(* IEC 61131-3 sources: Industry-PLC-LLM/data/PLCBEAD_repo/PLCBEAD_PLCEmbed-main/PLC-BEAD/Source/PLC_Programs (part 5) *)

(* ---- DT_TO_SDT.ST ---- *)
TYPE oscat_SDT :
STRUCT
	YEAR : INT;
	MONTH : INT;
	DAY : INT;
	WEEKDAY : INT;
	HOUR : INT;
	MINUTE : INT;
	SECOND : INT;
	MS : INT;
END_STRUCT;
END_TYPE

FUNCTION DT_TO_DATE2:UDINT

	VAR_INPUT
		IN :	UDINT;
	END_VAR

	DT_TO_DATE2 := (IN / UDINT#86400) * UDINT#86400;
END_FUNCTION

FUNCTION YEAR_OF_DATE:INT
	VAR_INPUT
		IDATE :	UDINT;
	END_VAR

	YEAR_OF_DATE := UDINT_TO_INT((idate+UDINT#43200) / UDINT#31557600 + UDINT#1970);
END_FUNCTION

FUNCTION DAY_OF_WEEK:INT

	VAR_INPUT
		IDATE :	UDINT;
	END_VAR

	DAY_OF_WEEK := UDINT_TO_INT((idate / UDINT#86400 + UDINT#3) MOD UDINT#7) + INT#01;
END_FUNCTION

FUNCTION LEAP_OF_DATE:BOOL

	VAR_INPUT
		IDATE :	UDINT;
	END_VAR

	LEAP_OF_DATE := SHL(UDINT_TO_DWORD((idate + UDINT#43200) / UDINT#31557600), 30) = DWORD#16#80000000;
END_FUNCTION

FUNCTION DAY_OF_YEAR:INT
	VAR_INPUT
		IDATE :	UDINT;
	END_VAR

	DAY_OF_YEAR := UDINT_TO_INT(((idate) / UDINT#86400) MOD UDINT#1461);
	IF DAY_OF_YEAR > 729 THEN
		IF DAY_OF_YEAR > 1095 THEN DAY_OF_YEAR := DAY_OF_YEAR - 1095; ELSE DAY_OF_YEAR := DAY_OF_YEAR - 729; END_IF;
	ELSIF DAY_OF_YEAR > 364 THEN
		DAY_OF_YEAR := DAY_OF_YEAR - 364;
	ELSE
		DAY_OF_YEAR := DAY_OF_YEAR + 1;
	END_IF;
END_FUNCTION

FUNCTION MONTH_OF_DATE:INT

	VAR_INPUT
		IDATE :	UDINT;
	END_VAR

	MONTH_OF_DATE := DAY_OF_YEAR(idate);
	IF MONTH_OF_DATE < 32 THEN
		MONTH_OF_DATE := 1;
	ELSIF LEAP_OF_DATE((IDATE)) THEN
		MONTH_OF_DATE := (MONTH_OF_DATE * 53 + 1668) / 1623;
	ELSE
		MONTH_OF_DATE := (MONTH_OF_DATE * 53 + 1700) / 1620;
	END_IF;
END_FUNCTION

FUNCTION DAY_OF_MONTH:INT
	VAR_INPUT
		IDATE :	UDINT;
	END_VAR

	day_of_month := day_of_year(idate);

	IF leap_of_Date((idate)) THEN
		CASE day_of_month OF
			32..60	:	day_of_month := day_of_month - 31;
			61..91	:	day_of_month := day_of_month - 60;
			92..121 :	day_of_month := day_of_month - 91;
			122..152:	day_of_month := day_of_month - 121;
			153..182:	day_of_month := day_of_month - 152;
			183..213:	day_of_month := day_of_month - 182;
			214..244:	day_of_month := day_of_month - 213;
			245..274:	day_of_month := day_of_month - 244;
			275..305:	day_of_month := day_of_month - 274;
			306..335:	day_of_month := day_of_month - 305;
			336..366:	day_of_month := day_of_month - 335;
		END_CASE;
	ELSE
		CASE day_of_month OF
			32..59	:	day_of_month := day_of_month - 31;
			60..90	:	day_of_month := day_of_month - 59;
			91..120 :	day_of_month := day_of_month - 90;
			121..151:	day_of_month := day_of_month - 120;
			152..181:	day_of_month := day_of_month - 151;
			182..212:	day_of_month := day_of_month - 181;
			213..243:	day_of_month := day_of_month - 212;
			244..273:	day_of_month := day_of_month - 243;
			274..304:	day_of_month := day_of_month - 273;
			305..334:	day_of_month := day_of_month - 304;
			335..365:	day_of_month := day_of_month - 334;
		END_CASE;
	END_IF;
END_FUNCTION

FUNCTION _INT_TO_UDINT:UDINT
	VAR_INPUT
		IN :	INT;
	END_VAR

	_INT_TO_UDINT := DINT_TO_UDINT(INT_TO_DINT(IN));
END_FUNCTION

FUNCTION_BLOCK DT_TO_SDT

	VAR_INPUT
		DTI :	UDINT;
	END_VAR

	VAR_OUTPUT
		SDT :	oscat_SDT;
	END_VAR

	VAR
		tmp :	UDINT;
		tdt :	UDINT;
	END_VAR

	tmp := DT_TO_DATE2(dti);
	tdt := dti - tmp;
	SDT.YEAR := YEAR_OF_DATE(tmp);
	SDT.MONTH := MONTH_OF_DATE(tmp);
	SDT.DAY := DAY_OF_MONTH(tmp);
	SDT.WEEKDAY := DAY_OF_WEEK(tmp);
	SDT.SECOND := UDINT_TO_INT(tdt MOD UDINT#60);
	SDT.MINUTE := UDINT_TO_INT((tdt / UDINT#60) MOD UDINT#60);
	SDT.HOUR := UDINT_TO_INT(tdt / UDINT#3600);

END_FUNCTION_BLOCK

PROGRAM program0
  VAR
    LocalVar0 : UDINT;
	LocalOUT  : oscat_SDT;
	func_block : DT_TO_SDT;
  END_VAR
	func_block.DTI  := LocalVar0;
	func_block();
	LocalOUT := func_block.SDT;
END_PROGRAM

CONFIGURATION Config0
  RESOURCE Res0 ON PLC
    TASK task0(INTERVAL := T#20ms,PRIORITY := 0);
    PROGRAM instance0 WITH task0 : program0;
  END_RESOURCE
END_CONFIGURATION

(* ---- DT_TO_STRF.ST ---- *)
FUNCTION DT_TO_DATE2:UDINT

	VAR_INPUT
		IN :	UDINT;
	END_VAR

	DT_TO_DATE2 := (IN / UDINT#86400) * UDINT#86400;
END_FUNCTION

FUNCTION DT_TO_TOD2:UDINT
	VAR_INPUT
		IN :	UDINT;
	END_VAR

	DT_TO_TOD2 := (IN MOD UDINT#86400) * UDINT#1000;
END_FUNCTION

FUNCTION _BYTE_TO_INT:INT
	VAR_INPUT
		IN :	BYTE;
	END_VAR

	_BYTE_TO_INT := USINT_TO_INT(BYTE_TO_USINT(IN));
END_FUNCTION

FUNCTION_BLOCK DT_TO_STRF_Block

	VAR_INPUT
		DTI :	UDINT;
		MS :	INT;
		FMT :	STRING;
		LANG :	INT;
	END_VAR

	VAR_OUTPUT
		DT_TO_STRF :	STRING;
	END_VAR

	VAR
		FILL :	STRING;
		BLANK :	STRING;
		ly :	INT;
		dx :	UDINT;
		fs :	STRING;
		fs_tmp :	STRING;
		td :	UDINT;
		tmp :	INT;
		pos :	INT;
		f :	INT;
		CODEE :	CODE;
		MONTH_TO_STRING :	MONTH_TO_STRING;
		WEEKDAY_TO_STRING :	WEEKDAY_TO_STRING;
	END_VAR

	IF LANG < 1 THEN ly := 1; ELSE ly := MIN(2, LANG); END_IF;

	dx := DT_TO_DATE2(DTI);
	td := DT_TO_TOD2(DTI);

	DT_TO_STRF := FMT;
	pos := FIND(DT_TO_STRF, '#');
	WHILE pos > 0 DO
		CODEE(STR:=DT_TO_STRF,POS:=pos + 1);
		f := _BYTE_TO_INT(CODEE.CODEE);
		(* generate the return string according to the format character *)
		fs := '';
		CASE f OF
			0: RETURN; (* illegal character index *)

			65 : (* letter A retunrs the year in 4 digits *)
				fs := INT_TO_STRING(YEAR_OF_DATE(dx),'%d');
			66 : (* letter B returns the year in exactly 2 digits *)
				fs := RIGHT(INT_TO_STRING(YEAR_OF_DATE(dx),'%02d'),2);
			67 : (* letter C returns the month with 1 or 2 digits *)
				fs := INT_TO_STRING(MONTH_OF_DATE(dx),'%d');
			68 : (* letter D returns the month with exactly 2 digits *)
				fs := INT_TO_STRING(MONTH_OF_DATE(dx),'%02d');
			69 : (* letter E returns the month with 3 characters *)
				MONTH_TO_STRING(MTH:=MONTH_OF_DATE(dx),LANG:=ly,LX:=3);
				fs:=MONTH_TO_STRING.MONTH_TO_STRING;
			70 : (* letter F returns the month with all characters *)
				MONTH_TO_STRING(MTH:=MONTH_OF_DATE(dx),LANG:=ly,LX:=0);
				fs:=MONTH_TO_STRING.MONTH_TO_STRING;
			71 : (* letter G returns the day with up to 2 digits *)
				fs := INT_TO_STRING(DAY_OF_MONTH(dx),'%d');
			72 : (* letter H returns the day of the month with exactly 2 digits *)
				fs := INT_TO_STRING(DAY_OF_MONTH(dx),'%d');
				IF LEN(fs) < 2 THEN fs_tmp:=fs; fs := CONCAT(FILL, fs_tmp); END_IF;
			73 : (* letter I returns the weekday as the number 1..7 1 = monday *)
				fs := INT_TO_STRING(DAY_OF_WEEK(dx),'%d');
			74 : (* letter J returns the weekday in 2 character writing *)
				WEEKDAY_TO_STRING(WDAY:=DAY_OF_WEEK(dx),LANG:=ly,LX:=2);
				fs := WEEKDAY_TO_STRING.WEEKDAY_TO_STRING;
			75 : (* letter K returns the weekday with all characters *)
				WEEKDAY_TO_STRING(WDAY:=DAY_OF_WEEK(dx),LANG:=ly,LX:=0);
				fs := WEEKDAY_TO_STRING.WEEKDAY_TO_STRING;
			76 : (* letter L returns AM or PM for the given DateTime *)
				IF td >= UDINT#43200000 THEN fs := 'PM'; ELSE fs := 'AM'; END_IF;
			77 : (* letter M returns the hour in 1 or 2 digit form 0..24h *)
				fs := INT_TO_STRING(HOUR(td),'%d');
			78 : (* letter N returns the hour in exactly 2 digit form 0..24h *)
				fs := INT_TO_STRING(HOUR(td),'%d');
				IF LEN(fs) < 2 THEN fs_tmp:=fs; fs := CONCAT(FILL, fs_tmp); END_IF;
			79 : (* letter O returns the hour in 1 or 2 digit form 0..12h *)
				tmp := HOUR(td) MOD 12;
				IF tmp = 0 THEN tmp := 12; END_IF;
				fs := INT_TO_STRING(tmp,'%d');
			80 : (* letter P returns the hour in exactly 2 digit form 0..12h *)
				tmp := HOUR(td) MOD 12;
				IF tmp = 0 THEN tmp := 12; END_IF;
				fs := INT_TO_STRING(tmp,'%d');
				IF LEN(fs) < 2 THEN fs_tmp:=fs; fs := CONCAT(FILL, fs_tmp); END_IF;
			81 : (* letter Q returns the minute of the hour in 1 or two digit form *)
				fs := INT_TO_STRING(MINUTE(td),'%d');
			82 : (* letter R returns the minute of the hour in exactly two digit form *)
				fs := INT_TO_STRING(MINUTE(td),'%d');
				IF LEN(fs) < 2 THEN fs_tmp:=fs; fs := CONCAT(FILL, fs_tmp); END_IF;
			83 : (* letter S returns the second of the minute in 1 or two digit form *)
				fs := INT_TO_STRING(REAL_TO_INT(SECOND(td)),'%d');
			84 : (* letter T returns the second of the minute in exactly two digit form *)
				fs := INT_TO_STRING(REAL_TO_INT(SECOND(td)),'%d');
				IF LEN(fs) < 2 THEN fs_tmp:=fs; fs := CONCAT(FILL, fs_tmp); END_IF;
			85 : (* letter U returns the milliseconds in 1 to 3 digits *)
				fs := INT_TO_STRING(MS,'%d');
			86 : (* letter V returns the milliseconds in exactly 3 digit form *)
				fs := INT_TO_STRING(MS,'%03d');
			87 : (* letter W returns the day of the month with exactly 2 digits first digit is filled with blank if necessary *)
				fs := INT_TO_STRING(DAY_OF_MONTH(dx),'%d');
				IF LEN(fs) < 2 THEN fs_tmp:=fs; fs := CONCAT(BLANK, fs_tmp); END_IF;
			88 : (* letter X returns the month with exactly 2 digits first digit is filled with blank if necessary *)
				fs := INT_TO_STRING(MONTH_OF_DATE(dx),'%d');
				IF LEN(fs) < 2 THEN fs_tmp:=fs; fs := CONCAT(BLANK, fs_tmp); END_IF;
		END_CASE;
		DT_TO_STRF := REPLACE(DT_TO_STRF, fs, 2, pos);
		pos := FIND(DT_TO_STRF, '#');
	END_WHILE;

END_FUNCTION_BLOCK

PROGRAM program0
  VAR
	DTI  :	UDINT;
	MS   :	INT;
	FMT  :	STRING;
	LANG :	INT;

	DT_TO_STRF :	STRING;

	func_block : DT_TO_STRF_Block;
  END_VAR
	func_block.DTI  :=DTI ;
	func_block.MS   :=MS  ;
	func_block.FMT  :=FMT ;
	func_block.LANG :=LANG;
	func_block();
	DT_TO_STRF := func_block.DT_TO_STRF;
END_PROGRAM

CONFIGURATION Config0
  RESOURCE Res0 ON PLC
    TASK task0(INTERVAL := T#20ms,PRIORITY := 0);
    PROGRAM instance0 WITH task0 : program0;
  END_RESOURCE
END_CONFIGURATION

(* ---- DT_TO_STRING.ST ---- *)
FUNCTION YEAR_OF_DATE:INT
	VAR_INPUT
		IDATE :	UDINT;
	END_VAR

	YEAR_OF_DATE := UDINT_TO_INT((idate+UDINT#43200) / UDINT#31557600 + UDINT#1970);
END_FUNCTION

FUNCTION DAY_OF_YEAR:INT
	VAR_INPUT
		IDATE :	UDINT;
	END_VAR

	DAY_OF_YEAR := UDINT_TO_INT(((idate) / UDINT#86400) MOD UDINT#1461);
	IF DAY_OF_YEAR > 729 THEN
		IF DAY_OF_YEAR > 1095 THEN DAY_OF_YEAR := DAY_OF_YEAR - 1095; ELSE DAY_OF_YEAR := DAY_OF_YEAR - 729; END_IF;
	ELSIF DAY_OF_YEAR > 364 THEN
		DAY_OF_YEAR := DAY_OF_YEAR - 364;
	ELSE
		DAY_OF_YEAR := DAY_OF_YEAR + 1;
	END_IF;
END_FUNCTION

FUNCTION LEAP_OF_DATE:BOOL

	VAR_INPUT
		IDATE :	UDINT;
	END_VAR

	LEAP_OF_DATE := SHL(UDINT_TO_DWORD((idate + UDINT#43200) / UDINT#31557600), 30) = DWORD#16#80000000;
END_FUNCTION

FUNCTION MONTH_OF_DATE:INT

	VAR_INPUT
		IDATE :	UDINT;
	END_VAR

	MONTH_OF_DATE := DAY_OF_YEAR(idate);
	IF MONTH_OF_DATE < 32 THEN
		MONTH_OF_DATE := 1;
	ELSIF LEAP_OF_DATE(IDATE) THEN
		MONTH_OF_DATE := (MONTH_OF_DATE * 53 + 1668) / 1623;
	ELSE
		MONTH_OF_DATE := (MONTH_OF_DATE * 53 + 1700) / 1620;
	END_IF;
END_FUNCTION

FUNCTION DAY_OF_MONTH:INT
	VAR_INPUT
		IDATE :	UDINT;
	END_VAR

	day_of_month := day_of_year(idate);

	IF leap_of_Date((idate)) THEN
		CASE day_of_month OF
			32..60	:	day_of_month := day_of_month - 31;
			61..91	:	day_of_month := day_of_month - 60;
			92..121 :	day_of_month := day_of_month - 91;
			122..152:	day_of_month := day_of_month - 121;
			153..182:	day_of_month := day_of_month - 152;
			183..213:	day_of_month := day_of_month - 182;
			214..244:	day_of_month := day_of_month - 213;
			245..274:	day_of_month := day_of_month - 244;
			275..305:	day_of_month := day_of_month - 274;
			306..335:	day_of_month := day_of_month - 305;
			336..366:	day_of_month := day_of_month - 335;
		END_CASE;
	ELSE
		CASE day_of_month OF
			32..59	:	day_of_month := day_of_month - 31;
			60..90	:	day_of_month := day_of_month - 59;
			91..120 :	day_of_month := day_of_month - 90;
			121..151:	day_of_month := day_of_month - 120;
			152..181:	day_of_month := day_of_month - 151;
			182..212:	day_of_month := day_of_month - 181;
			213..243:	day_of_month := day_of_month - 212;
			244..273:	day_of_month := day_of_month - 243;
			274..304:	day_of_month := day_of_month - 273;
			305..334:	day_of_month := day_of_month - 304;
			335..365:	day_of_month := day_of_month - 334;
		END_CASE;
	END_IF;
END_FUNCTION

FUNCTION SECOND_OF_DT:INT

	VAR_INPUT
		XDT :	UDINT;
	END_VAR

	SECOND_OF_DT := UDINT_TO_INT(XDT MOD UDINT#60);
END_FUNCTION

FUNCTION HOUR_OF_DT:INT
	VAR_INPUT
		XDT :	UDINT;
	END_VAR

	HOUR_OF_DT := UDINT_TO_INT((XDT MOD UDINT#86400) / UDINT#3600);
END_FUNCTION

FUNCTION MINUTE_OF_DT:INT
	VAR_INPUT
		XDT :	UDINT;
	END_VAR

	MINUTE_OF_DT := UDINT_TO_INT((XDT MOD UDINT#3600) / UDINT#60);
END_FUNCTION

FUNCTION_BLOCK DT_TO_STRING_Block

	VAR_INPUT
		IDT :	UDINT;
	END_VAR

	VAR_OUTPUT
		DT_STRING :	STRING;
	END_VAR

	VAR
		st_tmp1 :	STRING;
		st_tmp2 :	STRING;
	END_VAR

	st_tmp2 := CONCAT(INT_TO_STRING(YEAR_OF_DATE(IDT)),INT_TO_STRING(MONTH_OF_DATE(IDT)));
	st_tmp1 := CONCAT(INT_TO_STRING(day_of_month(IDT)),INT_TO_STRING(hour_of_DT(IDT)));
	st_tmp2 := CONCAT(st_tmp2,st_tmp1);
	st_tmp1 := CONCAT(INT_TO_STRING(minute_of_DT(IDT)),INT_TO_STRING(second_of_DT(IDT)));
	st_tmp2 := CONCAT(st_tmp2,st_tmp1);
	DT_STRING := st_tmp2;
END_FUNCTION_BLOCK

PROGRAM program0
	VAR
		IDT : UDINT;
		OUT  : STRING;
		func_block : DT_TO_STRING_Block;
	END_VAR
	func_block.IDT := IDT;
	func_block();
	OUT := func_block.DT_STRING;
END_PROGRAM

CONFIGURATION Config0
	RESOURCE Res0 ON PLC
		TASK task0(INTERVAL := T#20ms,PRIORITY := 0);
		PROGRAM instance0 WITH task0 : program0;
	END_RESOURCE
END_CONFIGURATION

(* ---- DW_TO_REAL.ST ---- *)
FUNCTION_BLOCK DW_TO_REAL_Block
  VAR_INPUT
    X :	DWORD;
  END_VAR

  VAR_OUTPUT
    DW_TO_REAL :	REAL;
  END_VAR

  VAR
    BUF_TO_REAL :	BUF_TO_REAL;
    i :	INT;
  END_VAR

  FOR I := 0 TO 1 DO
    BUF_TO_REAL.REQ        := I > 0;
    BUF_TO_REAL.BUF_FORMAT := FALSE;
    BUF_TO_REAL.BUF_OFFS   := DINT#0;
    BUF_TO_REAL.BUF_CNT    := DINT#4;
    BUF_TO_REAL.BUFFER     := X;
    BUF_TO_REAL.DST        := DW_TO_REAL;
    BUF_TO_REAL();
    X           := BUF_TO_REAL.BUFFER;
    DW_TO_REAL  := BUF_TO_REAL.DST;
  END_FOR;
END_FUNCTION_BLOCK

(* ---- DWORD_TO_STRB.ST ---- *)
FUNCTION_BLOCK DWORD_TO_STRB_Block
	VAR_INPUT
		IN :	DWORD;
	END_VAR

	VAR_OUTPUT
		DWORD_TO_STRB :	STRING;
	END_VAR

	VAR
		i :	INT;
	END_VAR

	DWORD_TO_STRB :='';
	FOR i := 1 TO 32 DO
		IF (in AND DWORD#16#8000_0000) > DWORD#0 THEN
			DWORD_TO_STRB := CONCAT(DWORD_TO_STRB,'1');
		ELSE
			DWORD_TO_STRB := CONCAT(DWORD_TO_STRB,'0');
		END_IF;
		in := SHL(in, 1);
	END_FOR;
END_FUNCTION_BLOCK

PROGRAM program0
  VAR
    IN :	DWORD;

	DWORD_TO_STRB :	STRING;
	func_block : DWORD_TO_STRB_Block;
  END_VAR
	func_block.IN  := IN;
	func_block();
	DWORD_TO_STRB := func_block.DWORD_TO_STRB;
END_PROGRAM

CONFIGURATION Config0
  RESOURCE Res0 ON PLC
    TASK task0(INTERVAL := T#20ms,PRIORITY := 0);
    PROGRAM instance0 WITH task0 : program0;
  END_RESOURCE
END_CONFIGURATION

(* ---- DWORD_TO_STRF.ST ---- *)
FUNCTION_BLOCK DWORD_TO_STRF_Block

	VAR_INPUT
		IN :	DWORD;
		N :	INT;
	END_VAR

	VAR_OUTPUT
		DWORD_TO_STRF :	STRING;
	END_VAR

	VAR
		temp :	STRING;
		temp2 :	STRING;
		L : INT;
	END_VAR

	temp := DWORD_TO_STRING(in);
	L := LEN(temp);
	IF N < L THEN
		temp :=RIGHT(temp,N);
		L := N;
	END_IF;

	WHILE L < N DO
		temp2 := temp;
		temp := CONCAT('0', temp2);
		L := L + 1;
	END_WHILE;
	DWORD_TO_STRF := temp;

END_FUNCTION_BLOCK

PROGRAM program0
  VAR
    IN :	DWORD;
	N :		INT;
	DWORD_TO_STRF :	STRING;
	func_block : DWORD_TO_STRF_Block;
  END_VAR
	func_block.IN  := IN;
	func_block.N  := N;
	func_block();
	DWORD_TO_STRF := func_block.DWORD_TO_STRF;
END_PROGRAM

CONFIGURATION Config0
  RESOURCE Res0 ON PLC
    TASK task0(INTERVAL := T#20ms,PRIORITY := 0);
    PROGRAM instance0 WITH task0 : program0;
  END_RESOURCE
END_CONFIGURATION

(* ---- DWORD_TO_STRH.ST ---- *)
FUNCTION_BLOCK DWORD_TO_STRH_Block

	VAR_INPUT
		IN :	DWORD;
	END_VAR

	VAR_OUTPUT
		DWORD_TO_STRH :	STRING;
	END_VAR

	DWORD_TO_STRH:=DWORD_TO_STRING(IN);

END_FUNCTION_BLOCK

PROGRAM program0
  VAR
    LocalVar0 : DWORD;
	LocalOUT  : STRING;
	func_block : DWORD_TO_STRH_Block;
  END_VAR
	func_block.IN  := LocalVar0;
	func_block();
	LocalOUT := func_block.DWORD_TO_STRH;
END_PROGRAM

CONFIGURATION Config0
  RESOURCE Res0 ON PLC
    TASK task0(INTERVAL := T#20ms,PRIORITY := 0);
    PROGRAM instance0 WITH task0 : program0;
  END_RESOURCE
END_CONFIGURATION

(* ---- ELEMENT_COUNT.ST ---- *)
TYPE
	oscat_STRING250             : STRING;
END_TYPE

FUNCTION_BLOCK ELEMENT_COUNT_Block

	VAR_IN_OUT
		ELEMENT :	oscat_STRING250;
	END_VAR

	VAR_INPUT
		SEP :	BYTE;
	END_VAR

	VAR_OUTPUT
		ELEMENT_COUNT :	INT;
	END_VAR

	VAR
		I :	INT;
		pos :	INT;
	END_VAR

	i := LEN(ELEMENT);
	IF i = 0 THEN
		ELEMENT_COUNT := 0;
	ELSE
		ELEMENT_COUNT := 1;
		FOR pos := 1 TO I DO
			IF INT_TO_BYTE(GET_CHAR(ELEMENT,pos)) = SEP THEN ELEMENT_COUNT := ELEMENT_COUNT + 1; END_IF;
		END_FOR;
	END_IF;

END_FUNCTION_BLOCK

PROGRAM program0
	VAR
		SEP :	BYTE;
		POS :	INT;
		ELEMENT :	oscat_STRING250;
		ELEMENT_GET :	oscat_STRING250;

		func_block : ELEMENT_COUNT_Block;
	END_VAR
	func_block.SEP    :=SEP    ;
	func_block.POS:=POS;
	func_block.ELEMENT     :=ELEMENT     ;
	func_block();
	ELEMENT    := func_block.ELEMENT    ;
	ELEMENT_GET:= func_block.ELEMENT_GET;

END_PROGRAM

CONFIGURATION Config0
  RESOURCE Res0 ON PLC
    TASK task0(INTERVAL := T#20ms,PRIORITY := 0);
    PROGRAM instance0 WITH task0 : program0;
  END_RESOURCE
END_CONFIGURATION

(* ---- ELEMENT_GET.ST ---- *)
TYPE
	oscat_STRING250             : STRING;
END_TYPE

FUNCTION_BLOCK ELEMENT_GET_Block

	VAR_INPUT
		SEP :	BYTE;
		POS :	INT;
	END_VAR

	VAR_IN_OUT
		ELEMENT :	oscat_STRING250;
	END_VAR

	VAR_OUTPUT
		ELEMENT_GET :	oscat_STRING250;
	END_VAR

	VAR
		i :	INT;
		i2 :	INT;
		cnt :	INT;
		size :	INT;
	END_VAR

	cnt := 0;
	size := LEN(ELEMENT);

	FOR i := 1 TO size DO
		IF cnt = POS THEN EXIT; END_IF;
		IF INT_TO_BYTE(GET_CHAR(ELEMENT,i)) = SEP THEN cnt := cnt + 1; END_IF;
	END_FOR;

	FOR i2 := i TO size DO
		IF INT_TO_BYTE(GET_CHAR(ELEMENT,i2)) = SEP THEN EXIT; END_IF;
	END_FOR;

	IF i2 > i THEN
		ELEMENT_GET := MID(ELEMENT,i2-i,i);
	ELSE
		ELEMENT_GET := '';
	END_IF;

END_FUNCTION_BLOCK

PROGRAM program0
	VAR
		SEP :	BYTE;
		POS :	INT;
		ELEMENT :	oscat_STRING250;
		ELEMENT_GET :	oscat_STRING250;

		func_block : ELEMENT_GET_Block;
	END_VAR
	func_block.SEP    :=SEP    ;
	func_block.POS:=POS;
	func_block.ELEMENT     :=ELEMENT     ;
	func_block();
	ELEMENT    := func_block.ELEMENT    ;
	ELEMENT_GET:= func_block.ELEMENT_GET;

END_PROGRAM

CONFIGURATION Config0
  RESOURCE Res0 ON PLC
    TASK task0(INTERVAL := T#20ms,PRIORITY := 0);
    PROGRAM instance0 WITH task0 : program0;
  END_RESOURCE
END_CONFIGURATION

(* ---- ENERGY.ST ---- *)
FUNCTION_BLOCK ENERGY
	VAR_INPUT
		J :	REAL;
		C :	REAL;
		WH :	REAL;
	END_VAR

	VAR_OUTPUT
		YJ :	REAL;
		YC :	REAL;
		YWH :	REAL;
	END_VAR

	YJ := J + Wh * 3600.0 + C * 4.1868;
	YC := YJ * 0.238845896627496;
	YWh := YJ * 2.7777777778E-004;
END_FUNCTION_BLOCK

PROGRAM program0
  VAR
		J  :	REAL;
		C  :	REAL;
		WH :	REAL;

		YJ  :	REAL;
		YC  :	REAL;
		YWH :	REAL;
	func_block : ENERGY;
  END_VAR
	func_block.J  :=J ;
	func_block.C  :=C ;
	func_block.WH :=WH;
	func_block();
	YJ  := func_block.YJ ;
	YC  := func_block.YC ;
	YWH := func_block.YWH;

END_PROGRAM

CONFIGURATION Config0
	RESOURCE Res0 ON PLC
		TASK task0(INTERVAL := T#20ms,PRIORITY := 0);
		PROGRAM instance0 WITH task0 : program0;
	END_RESOURCE
END_CONFIGURATION

(* ---- ESR_COLLECT.ST ---- *)
TYPE
	oscat_esr_collect_data      : ARRAY [0..7]    OF BYTE;
END_TYPE
TYPE oscat_esr_data :
  STRUCT
	typ    : BYTE;
	adress : STRING;
	DS     : UDINT;
	TS     : TIME;
	data   : oscat_esr_collect_data;
  END_STRUCT;
END_TYPE

TYPE
  oscat_ESR_3                : ARRAY [0..3] OF oscat_esr_data;
  oscat_ESR_31               : ARRAY [0..31] OF oscat_esr_data;
END_TYPE

FUNCTION INC1:INT

	VAR_INPUT
		X :	INT;
		N :	INT;
	END_VAR

	IF X >= N - 1 THEN
		INC1 := 0;
	ELSE
		INC1 := X + 1;
	END_IF;
END_FUNCTION

FUNCTION_BLOCK ESR_COLLECT
	VAR_INPUT
		ESR_0 :	oscat_ESR_3;
		ESR_1 :	oscat_ESR_3;
		ESR_2 :	oscat_ESR_3;
		ESR_3 :	oscat_ESR_3;
		ESR_4 :	oscat_ESR_3;
		ESR_5 :	oscat_ESR_3;
		ESR_6 :	oscat_ESR_3;
		ESR_7 :	oscat_ESR_3;
		RST :	BOOL;
	END_VAR

	VAR_IN_OUT
		POS :	INT;
	END_VAR

	VAR_OUTPUT
		ESR_OUT :	oscat_ESR_31;
	END_VAR

	VAR
		cnt :	INT := -1;
		max_in :	INT := 3;
		max_out :	INT := 32;
	END_VAR

	IF rst OR cnt < 0 THEN
		pos := -1;
	ELSE
		FOR cnt := 0 TO max_in DO
		IF esr_0[cnt].typ > BYTE#0 THEN pos := INC1(pos, max_out); esr_out[pos] := esr_0[cnt]; END_IF;
		IF esr_1[cnt].typ > BYTE#0 THEN pos := INC1(pos, max_out); esr_out[pos] := esr_1[cnt]; END_IF;
		IF esr_2[cnt].typ > BYTE#0 THEN pos := INC1(pos, max_out); esr_out[pos] := esr_2[cnt]; END_IF;
		IF esr_3[cnt].typ > BYTE#0 THEN pos := INC1(pos, max_out); esr_out[pos] := esr_3[cnt]; END_IF;
		IF esr_4[cnt].typ > BYTE#0 THEN pos := INC1(pos, max_out); esr_out[pos] := esr_4[cnt]; END_IF;
		IF esr_5[cnt].typ > BYTE#0 THEN pos := INC1(pos, max_out); esr_out[pos] := esr_5[cnt]; END_IF;
		IF esr_6[cnt].typ > BYTE#0 THEN pos := INC1(pos, max_out); esr_out[pos] := esr_6[cnt]; END_IF;
		IF esr_7[cnt].typ > BYTE#0 THEN pos := INC1(pos, max_out); esr_out[pos] := esr_7[cnt]; END_IF;
	END_FOR;
	END_IF;

END_FUNCTION_BLOCK

PROGRAM program0
  VAR
	ESR_0 :	oscat_ESR_3;
	ESR_1 :	oscat_ESR_3;
	ESR_2 :	oscat_ESR_3;
	ESR_3 :	oscat_ESR_3;
	ESR_4 :	oscat_ESR_3;
	ESR_5 :	oscat_ESR_3;
	ESR_6 :	oscat_ESR_3;
	ESR_7 :	oscat_ESR_3;
	RST   :	BOOL;

	POS   :	INT;

	ESR_OUT :	oscat_ESR_31;

	func_block : ESR_COLLECT;
  END_VAR
	func_block.ESR_0 :=ESR_0;
	func_block.ESR_1 :=ESR_1;
	func_block.ESR_2 :=ESR_2;
	func_block.ESR_3 :=ESR_3;
	func_block.ESR_4 :=ESR_4;
	func_block.ESR_5 :=ESR_5;
	func_block.ESR_6 :=ESR_6;
	func_block.ESR_7 :=ESR_7;
	func_block.RST   :=RST  ;
	func_block.POS   :=POS  ;

	func_block();
	POS := func_block.POS;
	ESR_OUT := func_block.ESR_OUT;

END_PROGRAM

CONFIGURATION Config0
	RESOURCE Res0 ON PLC
		TASK task0(INTERVAL := T#20ms,PRIORITY := 0);
		PROGRAM instance0 WITH task0 : program0;
	END_RESOURCE
END_CONFIGURATION

(* ---- ESR_MON_B8.ST ---- *)
TYPE
	oscat_esr_collect_data      : ARRAY [0..7]    OF BYTE;
END_TYPE
TYPE oscat_esr_data :
  STRUCT
	typ    : BYTE;
	adress : STRING;
	DS     : UDINT;
	TS     : TIME;
	data   : oscat_esr_collect_data;
  END_STRUCT;
END_TYPE

TYPE
  oscat_ESR_3                : ARRAY [0..3] OF oscat_esr_data;
  oscat_ESR_31               : ARRAY [0..31] OF oscat_esr_data;
END_TYPE

FUNCTION_BLOCK T_PLC_MS_block

	VAR_OUTPUT
		T_PLC_MS :	UDINT;
	END_VAR

	VAR_EXTERNAL
		PLC_TICKS_PER_SEC :	INT;
		PLC_SYS_TICK_CNT :	DINT;
	END_VAR

	VAR
		debug :	BOOL;(*Debug-Mode ON / OFF*)
		N :	INT;(*Debug-Faktor*)
		Offset :	UDINT;(*Debug-Offset*)
		temp :	DWORD := DWORD#1;(*Debug-Offset*)
		mode :	BOOL;(*modus*)
		faktor :	UDINT;(*Systemtakt-Faktor*)
		init :	BOOL;
		v_plc_ticks_per_sec :	UDINT;
		base :	UDINT := UDINT#1000;
	END_VAR

	IF init = FALSE THEN
		v_plc_ticks_per_sec := INT_TO_UDINT(PLC_TICKS_PER_SEC);
		IF v_plc_ticks_per_sec = UDINT#1024 THEN
			faktor := UDINT#1;
			mode := FALSE;
		ELSIF v_plc_ticks_per_sec > UDINT#0 THEN
			IF v_plc_ticks_per_sec <= base THEN
				faktor := base / v_plc_ticks_per_sec;
				mode := FALSE;
			ELSE
				faktor := v_plc_ticks_per_sec / base;
				mode := TRUE;
			END_IF;
		ELSE
			faktor := UDINT#1;
		END_IF;
		init := TRUE;
	END_IF;

	IF mode THEN
		T_PLC_MS := DINT_TO_UDINT(PLC_SYS_TICK_CNT) / faktor;
	ELSE
		T_PLC_MS := DINT_TO_UDINT(PLC_SYS_TICK_CNT) * faktor;
	END_IF;

	IF debug THEN
		T_PLC_MS := (DWORD_TO_UDINT(SHL(UDINT_TO_DWORD(T_PLC_MS),N) OR SHL(temp,N)) - UDINT#1) + Offset;
	END_IF;

END_FUNCTION_BLOCK

FUNCTION_BLOCK ESR_MON_B8

	VAR_INPUT
		S0 :	BOOL;
		A0 :	STRING;
		S1 :	BOOL;
		A1 :	STRING;
		S2 :	BOOL;
		A2 :	STRING;
		S3 :	BOOL;
		A3 :	STRING;
		S4 :	BOOL;
		A4 :	STRING;
		S5 :	BOOL;
		A5 :	STRING;
		S6 :	BOOL;
		A6 :	STRING;
		S7 :	BOOL;
		A7 :	STRING;
		DT_IN :	UDINT;
	END_VAR

	VAR_IN_OUT
		ESR_Out :	oscat_ESR_3;
	END_VAR

	VAR_OUTPUT
		ESR_FLAG :	BOOL;
	END_VAR

	VAR
		x0 :	BOOL;
		x1 :	BOOL;
		x2 :	BOOL;
		x3 :	BOOL;
		x4 :	BOOL;
		x5 :	BOOL;
		x6 :	BOOL;
		x7 :	BOOL;
		tx :	TIME;
		cnt :	INT;
		T_PLC_MS :	T_PLC_MS_block;
	END_VAR

	T_PLC_MS();
	tx:= UDINT_TO_TIME(T_PLC_MS.T_PLC_MS);

	ESR_Flag := FALSE;
	esr_out[3].typ := BYTE#0;
	esr_out[2].typ := BYTE#0;
	esr_out[1].typ := BYTE#0;
	esr_out[0].typ := BYTE#0;
	cnt := 0;

	IF s0 <> X0 THEN
		esr_out[cnt].typ := INT_TO_BYTE(10 + BOOL_TO_INT(s0));
		esr_out[cnt].adress := a0;
		esr_out[cnt].DS := DT_in;
		esr_out[cnt].TS := TX;
		X0 := S0;
		cnt := cnt + 1;
		esr_flag := TRUE;
	END_IF;
	IF s1 <> X1 THEN
		esr_out[cnt].typ := INT_TO_BYTE(10 + BOOL_TO_INT(s1));
		esr_out[cnt].adress := a1;
		esr_out[cnt].DS := DT_in;
		esr_out[cnt].TS := TX;
		X1 := S1;
		cnt := cnt + 1;
		esr_flag := TRUE;
	END_IF;
	IF s2 <> X2 THEN
		esr_out[cnt].typ := INT_TO_BYTE(10 + BOOL_TO_INT(s2));
		esr_out[cnt].adress := a2;
		esr_out[cnt].DS := DT_in;
		esr_out[cnt].TS := TX;
		X2 := S2;
		cnt := cnt + 1;
		esr_flag := TRUE;
	END_IF;
	IF s3 <> X3 THEN
		esr_out[cnt].typ := INT_TO_BYTE(10 + BOOL_TO_INT(s3));
		esr_out[cnt].adress := a3;
		esr_out[cnt].DS := DT_in;
		esr_out[cnt].TS := TX;
		X3 := S3;
		cnt := cnt + 1;
		esr_flag := TRUE;
	END_IF;
	IF s4 <> X4 AND cnt < 4 THEN
		esr_out[cnt].typ := INT_TO_BYTE(10 + BOOL_TO_INT(s4));
		esr_out[cnt].adress := a4;
		esr_out[cnt].DS := DT_in;
		esr_out[cnt].TS := TX;
		X4 := S4;
		cnt := cnt + 1;
		esr_flag := TRUE;
	END_IF;
	IF s5 <> X5  AND cnt < 4 THEN
		esr_out[cnt].typ := INT_TO_BYTE(10 + BOOL_TO_INT(s5));
		esr_out[cnt].adress := a5;
		esr_out[cnt].DS := DT_in;
		esr_out[cnt].TS := TX;
		X5 := S5;
		cnt := cnt + 1;
		esr_flag := TRUE;
	END_IF;
	IF s6 <> X6  AND cnt < 4 THEN
		esr_out[cnt].typ := INT_TO_BYTE(10 + BOOL_TO_INT(s6));
		esr_out[cnt].adress := a6;
		esr_out[cnt].DS := DT_in;
		esr_out[cnt].TS := TX;
		X6 := S6;
		cnt := cnt + 1;
		esr_flag := TRUE;
	END_IF;
	IF s7 <> X7  AND cnt < 4 THEN
		esr_out[cnt].typ := INT_TO_BYTE(10 + BOOL_TO_INT(s7));
		esr_out[cnt].adress := a7;
		esr_out[cnt].DS := DT_in;
		esr_out[cnt].TS := TX;
		X7 := S7;
		cnt := cnt + 1;
		esr_flag := TRUE;
	END_IF;

END_FUNCTION_BLOCK

PROGRAM program0

	VAR

		S0 :	BOOL;
		A0 :	STRING;
		S1 :	BOOL;
		A1 :	STRING;
		S2 :	BOOL;
		A2 :	STRING;
		S3 :	BOOL;
		A3 :	STRING;
		S4 :	BOOL;
		A4 :	STRING;
		S5 :	BOOL;
		A5 :	STRING;
		S6 :	BOOL;
		A6 :	STRING;
		S7 :	BOOL;
		A7 :	STRING;
		DT_IN   :	UDINT;

		ESR_Out :	oscat_ESR_3;

		ESR_FLAG :	BOOL;

		func_block : ESR_MON_B8;
  	END_VAR
	func_block.S0 := S0;
	func_block.A0 := A0;
	func_block.S1 := S1;
	func_block.A1 := A1;
	func_block.S2 := S2;
	func_block.A2 := A2;
	func_block.S3 := S3;
	func_block.A3 := A3;
	func_block.S4 := S4;
	func_block.A4 := A4;
	func_block.S5 := S5;
	func_block.A5 := A5;
	func_block.S6 := S6;
	func_block.A6 := A6;
	func_block.S7 := S7;
	func_block.A7 := A7;
	func_block.DT_IN := DT_IN;
	func_block.ESR_Out := ESR_Out;
	func_block();
	ESR_Out := func_block.ESR_Out;
	ESR_FLAG := func_block.ESR_FLAG;

END_PROGRAM

CONFIGURATION Config0

	VAR_GLOBAL
		PLC_TICKS_PER_SEC :	INT;
		PLC_SYS_TICK_CNT :	DINT;
	END_VAR

  	RESOURCE Res0 ON PLC
    	TASK task0(INTERVAL := T#20ms,PRIORITY := 0);
    	PROGRAM instance0 WITH task0 : program0;
  	END_RESOURCE

END_CONFIGURATION

(* ---- ESR_MON_R4.ST ---- *)
TYPE
	oscat_esr_collect_data      : ARRAY [0..7]    OF BYTE;
END_TYPE

TYPE oscat_esr_data :
  STRUCT
	typ    : BYTE;
	adress : STRING;
	DS     : UDINT;
	TS     : TIME;
	data   : oscat_esr_collect_data;
  END_STRUCT;
END_TYPE

TYPE
  oscat_ESR_3                : ARRAY [0..3] OF oscat_esr_data;
  oscat_ESR_31               : ARRAY [0..31] OF oscat_esr_data;
END_TYPE

FUNCTION_BLOCK REAL_TO_DW_Block
  VAR_INPUT
    X :	REAL;
  END_VAR

  VAR_OUTPUT
    REAL_TO_DW :	DWORD;
  END_VAR

  VAR
    REAL_TO_BUF :	REAL_TO_BUF;
    i :	INT;
  END_VAR

  FOR I := 0 TO 1 DO
    REAL_TO_BUF.REQ        := I > 0;
    REAL_TO_BUF.BUF_FORMAT := FALSE;
    REAL_TO_BUF.BUF_OFFS   := DINT#0;
    REAL_TO_BUF.BUF_CNT    := DINT#4;
    REAL_TO_BUF.SRC        := X;
    REAL_TO_BUF.BUFFER     := REAL_TO_DW;
    REAL_TO_BUF();
    X          := REAL_TO_BUF.SRC;
    REAL_TO_DW := REAL_TO_BUF.BUFFER;
  END_FOR;
END_FUNCTION_BLOCK

FUNCTION_BLOCK T_PLC_MS_block

	VAR_OUTPUT
		T_PLC_MS :	UDINT;
	END_VAR

	VAR_EXTERNAL
		PLC_TICKS_PER_SEC :	INT;
		PLC_SYS_TICK_CNT :	DINT;
	END_VAR

	VAR
		debug :	BOOL;(*Debug-Mode ON / OFF*)
		N :	INT;(*Debug-Faktor*)
		Offset :	UDINT;(*Debug-Offset*)
		temp :	DWORD := DWORD#1;(*Debug-Offset*)
		mode :	BOOL;(*modus*)
		faktor :	UDINT;(*Systemtakt-Faktor*)
		init :	BOOL;
		v_plc_ticks_per_sec :	UDINT;
		base :	UDINT := UDINT#1000;
	END_VAR

	IF init = FALSE THEN
		v_plc_ticks_per_sec := INT_TO_UDINT(PLC_TICKS_PER_SEC);
		IF v_plc_ticks_per_sec = UDINT#1024 THEN
			faktor := UDINT#1;
			mode := FALSE;
		ELSIF v_plc_ticks_per_sec > UDINT#0 THEN
			IF v_plc_ticks_per_sec <= base THEN
				faktor := base / v_plc_ticks_per_sec;
				mode := FALSE;
			ELSE
				faktor := v_plc_ticks_per_sec / base;
				mode := TRUE;
			END_IF;
		ELSE
			faktor := UDINT#1;
		END_IF;
		init := TRUE;
	END_IF;

	IF mode THEN
		T_PLC_MS := DINT_TO_UDINT(PLC_SYS_TICK_CNT) / faktor;
	ELSE
		T_PLC_MS := DINT_TO_UDINT(PLC_SYS_TICK_CNT) * faktor;
	END_IF;

	IF debug THEN
		T_PLC_MS := (DWORD_TO_UDINT(SHL(UDINT_TO_DWORD(T_PLC_MS),N) OR SHL(temp,N)) - UDINT#1) + Offset;
	END_IF;

END_FUNCTION_BLOCK

FUNCTION_BLOCK ESR_MON_R4
	VAR_INPUT
		R0 :	REAL;
		A0 :	STRING;
		S0 :	REAL;
		R1 :	REAL;
		A1 :	STRING;
		S1 :	REAL;
		R2 :	REAL;
		A2 :	STRING;
		S2 :	REAL;
		R3 :	REAL;
		A3 :	STRING;
		S3 :	REAL;
		DT_IN :	UDINT;
	END_VAR

	VAR_IN_OUT
		ESR_OUT :	oscat_ESR_3;
	END_VAR

	VAR_OUTPUT
		ESR_FLAG :	BOOL;
	END_VAR

	VAR
		x0 :	REAL;
		x1 :	REAL;
		x2 :	REAL;
		x3 :	REAL;
		tx :	TIME;
		cnt :	INT;
		T_PLC_MS :	T_PLC_MS_block;
		REAL_TO_DW :	REAL_TO_DW_Block;
		tmp :	DWORD;
	END_VAR

	T_PLC_MS();
	tx:= UDINT_TO_TIME(T_PLC_MS.T_PLC_MS);

	ESR_Flag := FALSE;
	esr_out[3].typ := BYTE#0;
	esr_out[2].typ := BYTE#0;
	esr_out[1].typ := BYTE#0;
	esr_out[0].typ := BYTE#0;
	cnt := 0;

	IF differ(R0, X0, S0) THEN
		REAL_TO_DW(X:=R0);
		tmp := REAL_TO_DW.REAL_TO_DW;

		esr_out[cnt].typ := BYTE#20;
		esr_out[cnt].adress := a0;
		esr_out[cnt].DS := DT_in;
		esr_out[cnt].TS := TX;
		esr_out[cnt].data[0] := Byte_of_Dword(tmp,BYTE#0);
		esr_out[cnt].data[1] := Byte_of_Dword(tmp,BYTE#1);
		esr_out[cnt].data[2] := Byte_of_Dword(tmp,BYTE#2);
		esr_out[cnt].data[3] := Byte_of_Dword(tmp,BYTE#3);
		X0 := R0;
		cnt := cnt + 1;
		esr_flag := TRUE;
	END_IF;
	IF differ(R1, X1, S1) THEN
		REAL_TO_DW(X:=R1);
		tmp := REAL_TO_DW.REAL_TO_DW;

		esr_out[cnt].typ := BYTE#20;
		esr_out[cnt].adress := a1;
		esr_out[cnt].DS := DT_in;
		esr_out[cnt].TS := TX;
		esr_out[cnt].data[0] := Byte_of_Dword(tmp,BYTE#0);
		esr_out[cnt].data[1] := Byte_of_Dword(tmp,BYTE#1);
		esr_out[cnt].data[2] := Byte_of_Dword(tmp,BYTE#2);
		esr_out[cnt].data[3] := Byte_of_Dword(tmp,BYTE#3);
		X1 := R1;
		cnt := cnt + 1;
		esr_flag := TRUE;
	END_IF;
	IF differ(R2, X2, S2) THEN
		REAL_TO_DW(X:=R2);
		tmp := REAL_TO_DW.REAL_TO_DW;

		esr_out[cnt].typ := BYTE#20;
		esr_out[cnt].adress := a2;
		esr_out[cnt].DS := DT_in;
		esr_out[cnt].TS := TX;
		esr_out[cnt].data[0] := Byte_of_Dword(tmp,BYTE#0);
		esr_out[cnt].data[1] := Byte_of_Dword(tmp,BYTE#1);
		esr_out[cnt].data[2] := Byte_of_Dword(tmp,BYTE#2);
		esr_out[cnt].data[3] := Byte_of_Dword(tmp,BYTE#3);
		X2 := R2;
		cnt := cnt + 1;
		esr_flag := TRUE;
	END_IF;
	IF differ(R3, X3, S3) THEN
		REAL_TO_DW(X:=R2);
		tmp := REAL_TO_DW.REAL_TO_DW;

		esr_out[cnt].typ := BYTE#20;
		esr_out[cnt].adress := a3;
		esr_out[cnt].DS := DT_in;
		esr_out[cnt].TS := TX;
		esr_out[cnt].data[0] := Byte_of_Dword(tmp,BYTE#0);
		esr_out[cnt].data[1] := Byte_of_Dword(tmp,BYTE#1);
		esr_out[cnt].data[2] := Byte_of_Dword(tmp,BYTE#2);
		esr_out[cnt].data[3] := Byte_of_Dword(tmp,BYTE#3);
		X3 := R3;
		cnt := cnt + 1;
		esr_flag := TRUE;
	END_IF;
END_FUNCTION_BLOCK

PROGRAM program0

	VAR
	VAR_INPUT
		R0 :	REAL;
		A0 :	STRING;
		S0 :	REAL;
		R1 :	REAL;
		A1 :	STRING;
		S1 :	REAL;
		R2 :	REAL;
		A2 :	STRING;
		S2 :	REAL;
		R3 :	REAL;
		A3 :	STRING;
		S3 :	REAL;
		DT_IN :	UDINT;

		ESR_OUT :	oscat_ESR_3;

		ESR_FLAG :	BOOL;

		func_block : ESR_MON_R4;
  	END_VAR
	func_block.R0 := R0;
	func_block.A0 := A0;
	func_block.S0 := S0;
	func_block.R1 := R1;
	func_block.A1 := A1;
	func_block.S1 := S1;
	func_block.R2 := R2;
	func_block.A2 := A2;
	func_block.S2 := S2;
	func_block.R3 := R3;
	func_block.A3 := A3;
	func_block.S3 := S3;
	func_block.DT_IN := DT_IN;
	func_block.ESR_Out := ESR_Out;
	func_block();
	ESR_Out := func_block.ESR_Out;
	ESR_FLAG := func_block.ESR_FLAG;

END_PROGRAM

CONFIGURATION Config0

	VAR_GLOBAL
		PLC_TICKS_PER_SEC :	INT;
		PLC_SYS_TICK_CNT :	DINT;
	END_VAR

  	RESOURCE Res0 ON PLC
    	TASK task0(INTERVAL := T#20ms,PRIORITY := 0);
    	PROGRAM instance0 WITH task0 : program0;
  	END_RESOURCE

END_CONFIGURATION

(* ---- ESR_MON_X8.ST ---- *)
TYPE
	oscat_esr_collect_data      : ARRAY [0..7]    OF BYTE;
END_TYPE

TYPE oscat_esr_data :
  STRUCT
	typ    : BYTE;
	adress : STRING;
	DS     : UDINT;
	TS     : TIME;
	data   : oscat_esr_collect_data;
  END_STRUCT;
END_TYPE

TYPE
  oscat_ESR_3                : ARRAY [0..3] OF oscat_esr_data;
  oscat_ESR_31               : ARRAY [0..31] OF oscat_esr_data;
END_TYPE

FUNCTION_BLOCK STATUS_TO_ESR_Block

	VAR_INPUT
		STATUS :	BYTE;
		ADRESS :	STRING;
		DT_IN :	UDINT;
		TS :	TIME;
	END_VAR

	VAR_OUTPUT
		STATUS_TO_ESR :	oscat_esr_data;
	END_VAR

	IF status < BYTE#100 THEN
		status_to_ESR.typ := BYTE#1;
	ELSIF status < BYTE#200 THEN
		status_to_ESR.typ := BYTE#2;
	ELSE
		status_to_ESR.typ := BYTE#3;
	END_IF;
	status_to_ESR.adress:= adress;
	status_to_ESR.DS := DT_in;
	status_to_ESR.TS := TS;
	status_to_ESR.data[0] := status;
END_FUNCTION_BLOCK

FUNCTION_BLOCK T_PLC_MS_block

	VAR_OUTPUT
		T_PLC_MS :	UDINT;
	END_VAR

	VAR_EXTERNAL
		PLC_TICKS_PER_SEC :	INT;
		PLC_SYS_TICK_CNT :	DINT;
	END_VAR

	VAR
		debug :	BOOL;(*Debug-Mode ON / OFF*)
		N :	INT;(*Debug-Faktor*)
		Offset :	UDINT;(*Debug-Offset*)
		temp :	DWORD := DWORD#1;(*Debug-Offset*)
		mode :	BOOL;(*modus*)
		faktor :	UDINT;(*Systemtakt-Faktor*)
		init :	BOOL;
		v_plc_ticks_per_sec :	UDINT;
		base :	UDINT := UDINT#1000;
	END_VAR

	IF init = FALSE THEN
		v_plc_ticks_per_sec := INT_TO_UDINT(PLC_TICKS_PER_SEC);
		IF v_plc_ticks_per_sec = UDINT#1024 THEN
			faktor := UDINT#1;
			mode := FALSE;
		ELSIF v_plc_ticks_per_sec > UDINT#0 THEN
			IF v_plc_ticks_per_sec <= base THEN
				faktor := base / v_plc_ticks_per_sec;
				mode := FALSE;
			ELSE
				faktor := v_plc_ticks_per_sec / base;
				mode := TRUE;
			END_IF;
		ELSE
			faktor := UDINT#1;
		END_IF;
		init := TRUE;
	END_IF;

	IF mode THEN
		T_PLC_MS := DINT_TO_UDINT(PLC_SYS_TICK_CNT) / faktor;
	ELSE
		T_PLC_MS := DINT_TO_UDINT(PLC_SYS_TICK_CNT) * faktor;
	END_IF;

	IF debug THEN
		T_PLC_MS := (DWORD_TO_UDINT(SHL(UDINT_TO_DWORD(T_PLC_MS),N) OR SHL(temp,N)) - UDINT#1) + Offset;
	END_IF;

END_FUNCTION_BLOCK

FUNCTION_BLOCK ESR_MON_X8
	VAR_INPUT
		S0 :	BYTE;
		A0 :	STRING;
		S1 :	BYTE;
		A1 :	STRING;
		S2 :	BYTE;
		A2 :	STRING;
		S3 :	BYTE;
		A3 :	STRING;
		S4 :	BYTE;
		A4 :	STRING;
		S5 :	BYTE;
		A5 :	STRING;
		S6 :	BYTE;
		A6 :	STRING;
		S7 :	BYTE;
		A7 :	STRING;
		DT_IN :	UDINT;
		MODE :	BYTE := BYTE#3;
	END_VAR

	VAR_IN_OUT
		ESR_OUT :	oscat_ESR_3;
	END_VAR

	VAR_OUTPUT
		ESR_FLAG :	BOOL;
	END_VAR

	VAR
		x0 :	BYTE;
		x1 :	BYTE;
		x2 :	BYTE;
		x3 :	BYTE;
		x4 :	BYTE;
		x5 :	BYTE;
		x6 :	BYTE;
		x7 :	BYTE;
		tx :	TIME;
		cnt :	INT;
		status_to_ESR :	STATUS_TO_ESR_Block;
		T_PLC_MS :	T_PLC_MS_block;
	END_VAR

	T_PLC_MS();
	tx:= UDINT_TO_TIME(T_PLC_MS.T_PLC_MS);

	ESR_Flag := FALSE;
	esr_out[3].typ := BYTE#0;
	esr_out[2].typ := BYTE#0;
	esr_out[1].typ := BYTE#0;
	esr_out[0].typ := BYTE#0;
	cnt := 0;

	IF s0 <> X0 AND ((s0 < BYTE#100) OR (S0 > BYTE#99 AND S0 < BYTE#200 AND mode >= BYTE#2) OR (S0 > BYTE#199 AND mode = BYTE#3)) THEN

		status_to_ESR.status := s0;
		status_to_ESR.adress := a0;
		status_to_ESR.DT_in  := DT_in;
		status_to_ESR.TS     := tx;
		status_to_ESR();
		esr_out[cnt] := status_to_ESR.status_to_ESR;

		X0 := S0;
		cnt := cnt + 1;
		esr_flag := TRUE;
	END_IF;
	IF s1 <> X1 AND ((s1 < BYTE#100) OR (S1 > BYTE#99 AND S1 < BYTE#200 AND mode >= BYTE#2) OR (S1 > BYTE#199 AND mode = BYTE#3)) THEN

		status_to_ESR.status := s1;
		status_to_ESR.adress := a1;
		status_to_ESR.DT_in  := DT_in;
		status_to_ESR.TS     := tx;
		status_to_ESR();
		esr_out[cnt] := status_to_ESR.status_to_ESR;

		X1 := S1;
		cnt := cnt + 1;
		esr_flag := TRUE;
	END_IF;
	IF s2 <> X2 AND ((s2 < BYTE#100) OR (S2 > BYTE#99 AND S2 < BYTE#200 AND mode >= BYTE#2) OR (S2 > BYTE#199 AND mode = BYTE#3)) THEN

		status_to_ESR.status := s2;
		status_to_ESR.adress := a2;
		status_to_ESR.DT_in  := DT_in;
		status_to_ESR.TS     := tx;
		status_to_ESR();
		esr_out[cnt] := status_to_ESR.status_to_ESR;

		X2 := S2;
		cnt := cnt + 1;
		esr_flag := TRUE;
	END_IF;
	IF s3 <> X3 AND ((s3 < BYTE#100) OR (S3 > BYTE#99 AND S3 < BYTE#200 AND mode >= BYTE#2) OR (S3 > BYTE#199 AND mode = BYTE#3)) THEN

		status_to_ESR.status := s3;
		status_to_ESR.adress := a3;
		status_to_ESR.DT_in  := DT_in;
		status_to_ESR.TS     := tx;
		status_to_ESR();
		esr_out[cnt] := status_to_ESR.status_to_ESR;

		X3 := S3;
		cnt := cnt + 1;
		esr_flag := TRUE;
	END_IF;
	IF cnt < 4 AND s4 <> X4 AND ((s4 < BYTE#100) OR (S4 > BYTE#99 AND S4 < BYTE#200 AND mode >= BYTE#2) OR (S4 > BYTE#199 AND mode = BYTE#3)) THEN

		status_to_ESR.status := s4;
		status_to_ESR.adress := a4;
		status_to_ESR.DT_in  := DT_in;
		status_to_ESR.TS     := tx;
		status_to_ESR();
		esr_out[cnt] := status_to_ESR.status_to_ESR;

		X4 := S4;
		cnt := cnt + 1;
		esr_flag := TRUE;
	END_IF;
	IF cnt < 4 AND s5 <> X5 AND ((s5 < BYTE#100) OR (S5 > BYTE#99 AND S5 < BYTE#200 AND mode >= BYTE#2) OR (S5 > BYTE#199 AND mode = BYTE#3)) THEN

		status_to_ESR.status := s5;
		status_to_ESR.adress := a5;
		status_to_ESR.DT_in  := DT_in;
		status_to_ESR.TS     := tx;
		status_to_ESR();
		esr_out[cnt] := status_to_ESR.status_to_ESR;

		X5 := S5;
		cnt := cnt + 1;
		esr_flag := TRUE;
	END_IF;
	IF cnt < 4 AND s6 <> X6 AND ((s6 < BYTE#100) OR (S6 > BYTE#99 AND S6 < BYTE#200 AND mode >= BYTE#2) OR (S6 > BYTE#199 AND mode = BYTE#3)) THEN

		status_to_ESR.status := s6;
		status_to_ESR.adress := a6;
		status_to_ESR.DT_in  := DT_in;
		status_to_ESR.TS     := tx;
		status_to_ESR();
		esr_out[cnt] := status_to_ESR.status_to_ESR;

		X6 := S6;
		cnt := cnt + 1;
		esr_flag := TRUE;
	END_IF;
	IF cnt < 4 AND s7 <> X7 AND ((s7 < BYTE#100) OR (S7 > BYTE#99 AND S7 < BYTE#200 AND mode >= BYTE#2) OR (S7 > BYTE#199 AND mode = BYTE#3)) THEN

		status_to_ESR.status := s7;
		status_to_ESR.adress := a7;
		status_to_ESR.DT_in  := DT_in;
		status_to_ESR.TS     := tx;
		status_to_ESR();
		esr_out[cnt] := status_to_ESR.status_to_ESR;

		X7 := S7;
		cnt := cnt + 1;
		esr_flag := TRUE;
	END_IF;

END_FUNCTION_BLOCK

PROGRAM program0

	VAR
	S0 :	BYTE;
	A0 :	STRING;
	S1 :	BYTE;
	A1 :	STRING;
	S2 :	BYTE;
	A2 :	STRING;
	S3 :	BYTE;
	A3 :	STRING;
	S4 :	BYTE;
	A4 :	STRING;
	S5 :	BYTE;
	A5 :	STRING;
	S6 :	BYTE;
	A6 :	STRING;
	S7 :	BYTE;
	A7 :	STRING;
	DT_IN :	UDINT;
	MODE :	BYTE;

	ESR_OUT :	oscat_ESR_3;

	ESR_FLAG :	BOOL;

		func_block : ESR_MON_X8;
  	END_VAR
	func_block.S0 := S0;
	func_block.A0 := A0;
	func_block.S1 := S1;
	func_block.A1 := A1;
	func_block.S2 := S2;
	func_block.A2 := A2;
	func_block.S3 := S3;
	func_block.A3 := A3;
	func_block.S4 := S4;
	func_block.A4 := A4;
	func_block.S5 := S5;
	func_block.A5 := A5;
	func_block.S6 := S6;
	func_block.A6 := A6;
	func_block.S7 := S7;
	func_block.A7 := A7;
	func_block.DT_IN := DT_IN;
	func_block.MODE := MODE;
	func_block.ESR_Out := ESR_Out;
	func_block();
	ESR_Out := func_block.ESR_Out;
	ESR_FLAG := func_block.ESR_FLAG;
END_PROGRAM

CONFIGURATION Config0

	VAR_GLOBAL
		PLC_TICKS_PER_SEC :	INT;
		PLC_SYS_TICK_CNT :	DINT;
	END_VAR

  	RESOURCE Res0 ON PLC
    	TASK task0(INTERVAL := T#20ms,PRIORITY := 0);
    	PROGRAM instance0 WITH task0 : program0;
  	END_RESOURCE

END_CONFIGURATION

(* ---- EVENTS.ST ---- *)
TYPE oscat_HOLIDAY_DATA :
  STRUCT
	NAME : STRING;
	DAY : SINT;
	MONTH : SINT;
	USE : SINT;
	PAD_BYTE : BYTE;
  END_STRUCT;
END_TYPE

TYPE
  oscat_HOLIDAY_DATA_0_29 	: ARRAY [0..29] OF oscat_HOLIDAY_DATA;
  oscat_HOLIDAY_DATA_0_49 	: ARRAY [0..49] OF oscat_HOLIDAY_DATA;
END_TYPE

FUNCTION DAY_OF_DATE:DINT
	VAR_INPUT
		IDATE :	UDINT;
	END_VAR

	day_of_date := UDINT_TO_DINT(idate / UDINT#86400);
END_FUNCTION

FUNCTION YEAR_OF_DATE:INT
	VAR_INPUT
		IDATE :	UDINT;
	END_VAR

	YEAR_OF_DATE := UDINT_TO_INT((idate+UDINT#43200) / UDINT#31557600 + UDINT#1970);
END_FUNCTION

FUNCTION _INT_TO_UDINT:UDINT
	VAR_INPUT
		IN :	INT;
	END_VAR

	_INT_TO_UDINT := DINT_TO_UDINT(INT_TO_DINT(IN));
END_FUNCTION

FUNCTION SET_DATE:UDINT

	VAR_INPUT
		YEAR :	INT;
		MONTH :	INT;
		DAY :	INT;
	END_VAR

	VAR
		count :	INT;
	END_VAR

	IF month > 2 THEN
		count := (month - 1) * 30;
		IF month > 7 THEN
			count := count + DWORD_TO_INT(SHR(DINT_TO_DWORD(INT_TO_DINT(month) - INT_TO_DINT(3)),1));
		ELSE
			count := count + DWORD_TO_INT(SHR(DINT_TO_DWORD(INT_TO_DINT(month) - INT_TO_DINT(4)),1));
		END_IF;
		IF SHL(INT_TO_WORD(year),14) = WORD#0 THEN
			count := count + 1;
		END_IF;
	ELSE
		count := (month - 1) * 31;
	END_IF;
	SET_DATE := (_INT_TO_UDINT(count + day - 1) + DWORD_TO_UDINT(SHR(UDINT_TO_DWORD(_INT_TO_UDINT(year) * UDINT#1461 - UDINT#2878169), 2))) * UDINT#86400;
END_FUNCTION

FUNCTION_BLOCK EVENTS
	VAR_INPUT
		DATE_IN :	UDINT;
		ENA :	BOOL;
	END_VAR

	VAR_OUTPUT
		Y :	BOOL;
		NAME :	STRING;
	END_VAR

	VAR_IN_OUT
		ELIST :	oscat_HOLIDAY_DATA_0_49;
	END_VAR

	VAR
		i :	INT;
		last_active :	UDINT;
		size :	INT := 49;
		day_in :	DINT;
		cyr :	INT;
		lday :	DINT;
		check :	oscat_HOLIDAY_DATA;
		y_int :	BOOL;
		name_int :	STRING;
	END_VAR

	IF last_active <> date_in THEN
		last_active := DATE_IN;
		Y_int := FALSE;
		name_int := '';
		day_in := DAY_OF_DATE(DATE_IN);
		cyr := YEAR_OF_DATE(DATE_IN);

		(* search list for events *)
		FOR i := 0 TO size DO
			check := elist[i];
			lday := DAY_OF_DATE(SET_DATE(cyr,SINT_TO_INT(check.month), SINT_TO_INT(check.day)));
			IF day_in >= lday AND day_in <= lday + SINT_TO_DINT(check.use) - DINT#1 THEN
				y_int := TRUE;
				name_int := check.name;
				EXIT;
			END_IF;
		END_FOR;
	END_IF;

	IF ENA THEN
		Y := y_int;
		NAME := name_int;
	ELSE
		Y := FALSE;
		NAME := '';
	END_IF;

END_FUNCTION_BLOCK

PROGRAM program0
	VAR
		DATE_IN :	UDINT;
		ENA :	BOOL;

		Y :	BOOL;
		NAME :	STRING;

		ELIST :	oscat_HOLIDAY_DATA_0_49;

		func_block : EVENTS;
	END_VAR
	func_block.DATE_IN := DATE_IN;
	func_block.ENA := ENA;
	func_block.ELIST := ELIST ;

	func_block();
	Y  := func_block.Y;
	NAME  := func_block.NAME;
	ELIST  := func_block.ELIST;
END_PROGRAM

CONFIGURATION Config0
	RESOURCE Res0 ON PLC
		TASK task0(INTERVAL := T#20ms,PRIORITY := 0);
		PROGRAM instance0 WITH task0 : program0;
	END_RESOURCE
END_CONFIGURATION

(* ---- EXEC.ST ---- *)
FUNCTION_BLOCK EXEC_Block
	VAR_INPUT
		STR :	STRING;
	END_VAR

	VAR_OUTPUT
		EXEC :	STRING;
	END_VAR

	VAR
		pos :	INT;
		R1 :	REAL;
		R2 :	REAL;
		operator :	STRING;
		temp :	STRING;
		uppercase :	uppercase;
		trim :	trim;
		findB_num :	findB_num;
		findB_nonum :	findB_nonum;
	END_VAR

	trim(str:=str);
	temp:=trim.trim;

	uppercase(str:=temp);
	exec:=uppercase.uppercase;

	findB_nonum(str:=exec);
	pos :=findB_nonum.findB_nonum;

	IF pos > 1 THEN
	temp := LEFT(EXEC,pos-1);
	findB_num(str:=temp);
	IF findB_num.findB_num > 0 THEN
	R1 := STRING_TO_REAL(temp);
	END_IF;
	END_IF;
	temp := RIGHT(exec,LEN(exec)-pos);
	R2 := STRING_TO_REAL(temp);
	exec := LEFT(exec,pos);

	findB_num(str:=exec);
	pos :=findB_num.findB_num;
	operator := RIGHT(exec,LEN(exec) - pos);
	IF EQ_STRING(operator,'') AND LEN(str) = 0 THEN
		exec := '';
		RETURN;
	ELSIF EQ_STRING(operator,'') THEN
		exec := str;
		RETURN;
	END_IF;
	IF EQ_STRING(operator,'^') THEN
		exec := REAL_TO_STRING(EXPT(R1, R2),'%f');
	ELSIF EQ_STRING(operator,'SQRT') THEN
		exec := REAL_TO_STRING(SQRT(R2),'%f');
	ELSIF EQ_STRING(operator,'SIN') THEN
		exec := REAL_TO_STRING(SIN(r2),'%f');
	ELSIF EQ_STRING(operator,'COS') THEN
		exec := REAL_TO_STRING(COS(r2),'%f');
	ELSIF EQ_STRING(operator,'TAN') THEN
		exec := REAL_TO_STRING(TAN(R2),'%f');
	ELSIF EQ_STRING(operator,'*') THEN
		exec := REAL_TO_STRING(R1 * R2,'%f');
	ELSIF EQ_STRING(operator,'/') THEN
		IF R2 <> 0.0 THEN exec := REAL_TO_STRING(R1 / R2,'%f'); ELSE exec := 'ERROR'; END_IF;
	ELSIF EQ_STRING(operator,'+') THEN
		exec := REAL_TO_STRING(r1 + r2,'%f');
	ELSIF EQ_STRING(operator,'-') THEN
		exec := REAL_TO_STRING(r1 - r2,'%f');
	ELSE
		exec := 'ERROR';
	END_IF;
	IF EQ_STRING(EXEC,'ERROR') THEN
		RETURN;
	ELSIF FIND(EXEC,'.') = 0 THEN
		EXEC := CONCAT(EXEC, '.0');
	ELSE
	temp := RIGHT(EXEC,1);
	IF EQ_STRING(temp,'.') THEN
		EXEC := CONCAT(EXEC,'0');
	END_IF;
	END_IF;

END_FUNCTION_BLOCK

PROGRAM program0
	VAR
		STR :	STRING;

		EXEC :	STRING;

		func_block : EXEC_Block;
	END_VAR
	func_block.STR := STR;
	func_block();
	EXEC  := func_block.EXEC;
END_PROGRAM

CONFIGURATION Config0
	RESOURCE Res0 ON PLC
		TASK task0(INTERVAL := T#20ms,PRIORITY := 0);
		PROGRAM instance0 WITH task0 : program0;
	END_RESOURCE
END_CONFIGURATION

(* ---- F_LAMP.ST ---- *)
FUNCTION_BLOCK T_PLC_MS_block
	VAR_OUTPUT
		T_PLC_MS :	UDINT;
	END_VAR

	VAR_EXTERNAL
		PLC_TICKS_PER_SEC :	INT;
		PLC_SYS_TICK_CNT :	DINT;
	END_VAR

	VAR
		debug :	BOOL;(*Debug-Mode ON / OFF*)
		N :	INT;(*Debug-Faktor*)
		Offset :	UDINT;(*Debug-Offset*)
		temp :	DWORD := DWORD#1;(*Debug-Offset*)
		mode :	BOOL;(*modus*)
		faktor :	UDINT;(*Systemtakt-Faktor*)
		init :	BOOL;
		v_plc_ticks_per_sec :	UDINT;
		base :	UDINT := UDINT#1000;
	END_VAR

	IF init = FALSE THEN
		v_plc_ticks_per_sec := INT_TO_UDINT(PLC_TICKS_PER_SEC);
		IF v_plc_ticks_per_sec = UDINT#1024 THEN
			faktor := UDINT#1;
			mode := FALSE;
		ELSIF v_plc_ticks_per_sec > UDINT#0 THEN
			IF v_plc_ticks_per_sec <= base THEN
				faktor := base / v_plc_ticks_per_sec;
				mode := FALSE;
			ELSE
				faktor := v_plc_ticks_per_sec / base;
				mode := TRUE;
			END_IF;
		ELSE
			faktor := UDINT#1;
		END_IF;
		init := TRUE;
	END_IF;

	IF mode THEN
		T_PLC_MS := DINT_TO_UDINT(PLC_SYS_TICK_CNT) / faktor;
	ELSE
		T_PLC_MS := DINT_TO_UDINT(PLC_SYS_TICK_CNT) * faktor;
	END_IF;

	IF debug THEN
		T_PLC_MS := (DWORD_TO_UDINT(SHL(UDINT_TO_DWORD(T_PLC_MS),N) OR SHL(temp,N)) - UDINT#1) + Offset;
	END_IF;

END_FUNCTION_BLOCK

FUNCTION_BLOCK ONTIME_Block

	VAR_INPUT
		IN :	BOOL;
		RST :	BOOL;
	END_VAR

	VAR_IN_OUT
		SECONDS :	UDINT;
		CYCLES :	UDINT;
	END_VAR

	VAR
		tx :	UDINT;
		last :	UDINT;
		edge :	BOOL;
		init :	BOOL;
		ms :	UDINT;
		T_PLC_MS :	T_PLC_MS_Block;
	END_VAR

	T_PLC_MS();
	tx:= T_PLC_MS.T_PLC_MS;

	IF NOT init THEN
		init := TRUE;
		last := tx;
		ms := UDINT#0;
	END_IF;
	IF RST THEN
		SECONDS := UDINT#0;
		CYCLES := UDINT#0;
		last := tx;
		ms := UDINT#0;
	ELSIF IN THEN
		(* add the current milliseconds *)
		ms := (tx - last) + ms;
		IF ms >= UDINT#1000 THEN
			seconds := seconds + UDINT#1;
			ms := ms - UDINT#1000;
		END_IF;
		cycles := cycles + BOOL_TO_UDINT(NOT edge);
	END_IF;
	last := tx;
	edge := in;

END_FUNCTION_BLOCK

FUNCTION_BLOCK F_LAMP_Block

	VAR_INPUT
		SWITCH :	BOOL;
		DIMM :	BYTE := BYTE#255;
		RST :	BOOL;
		T_NO_DIMM :	UINT := UINT#100;
		T_MAINTENANCE :	UINT := UINT#15000;
	END_VAR

	VAR_OUTPUT
		LAMP :	BYTE;
		STATUS :	BYTE;
	END_VAR

	VAR_IN_OUT
		ONTIME :	UDINT;
		CYCLES :	UDINT;
	END_VAR

	VAR
		runtime :	ONTIME_Block;
	END_VAR

	runtime(in := switch, SECONDS := ONTIME , CYCLES := CYCLES);
	CYCLES := runtime.CYCLES;
	ONTIME := runtime.SECONDS;

	IF RST THEN
		ONTIME := UDINT#0;
		CYCLES := UDINT#0;
	END_IF;
	IF SWITCH THEN
		IF ontime < UINT_TO_UDINT(T_NO_DIMM) * UDINT#3600 THEN
			LAMP := BYTE#255;
			STATUS := BYTE#111;
		ELSE
			LAMP := DIMM;
			STATUS := BYTE#112;
		END_IF;
	ELSE
		LAMP := BYTE#0;
		STATUS := BYTE#110;
	END_IF;

	IF ontime >= UINT_TO_UDINT(T_maintenance) * UDINT#3600 AND T_Maintenance > UINT#0 THEN
		STATUS := BYTE#120;
	END_IF;

END_FUNCTION_BLOCK

PROGRAM program0
	VAR
	    SWITCH :	BOOL;
		DIMM :	BYTE := BYTE#255;
		RST :	BOOL;
		T_NO_DIMM :	UINT := UINT#100;
		T_MAINTENANCE :	UINT := UINT#15000;
		ONTIME :	UDINT;
		CYCLES :	UDINT;
		LAMP :	BYTE;
		STATUS :	BYTE;

		func_block : F_LAMP_Block;
  	END_VAR
	func_block.SWITCH := SWITCH;
	func_block.DIMM := DIMM;
	func_block.RST := RST;
	func_block.T_NO_DIMM := T_NO_DIMM;
	func_block.T_MAINTENANCE := T_MAINTENANCE;
	func_block.ONTIME := ONTIME;
	func_block.CYCLES := CYCLES;

	func_block();
	ONTIME := func_block.ONTIME;
	CYCLES := func_block.CYCLES;
	LAMP := func_block.LAMP;
	STATUS := func_block.STATUS;
END_PROGRAM

CONFIGURATION Config0
	VAR_GLOBAL
		PLC_TICKS_PER_SEC :	INT;
		PLC_SYS_TICK_CNT :	DINT;
	END_VAR
  	RESOURCE Res0 ON PLC
    	TASK task0(INTERVAL := T#20ms,PRIORITY := 0);
    	PROGRAM instance0 WITH task0 : program0;
  	END_RESOURCE
END_CONFIGURATION

(* ---- F_POLY.ST ---- *)
TYPE
  oscat_arr_0_7               : ARRAY [0..7]    OF REAL;
END_TYPE

FUNCTION_BLOCK F_POLY_Block
	VAR_INPUT
		X :	REAL;
		C :	oscat_arr_0_7;
	END_VAR

	VAR_OUTPUT
		F_POLY :	REAL;
	END_VAR

	F_POLY := ((((((( c[7] * x + c[6] ) * x + c[5] ) * x + c[4] ) * x + c[3] ) * x + c[2] ) * x + c[1] ) * x + c[0] ) ;

END_FUNCTION_BLOCK

PROGRAM program0
	VAR
		X :	REAL;
		C :	oscat_arr_0_7;

		F_POLY :	REAL;

		func_block : F_POLY_Block;
	END_VAR
	func_block.X := X;
	func_block.C := C;
	func_block();
	F_POLY  := func_block.F_POLY;
END_PROGRAM

CONFIGURATION Config0
	RESOURCE Res0 ON PLC
		TASK task0(INTERVAL := T#20ms,PRIORITY := 0);
		PROGRAM instance0 WITH task0 : program0;
	END_RESOURCE
END_CONFIGURATION

(* ---- FADE.ST ---- *)
FUNCTION_BLOCK T_PLC_MS_block
	VAR_OUTPUT
		T_PLC_MS :	UDINT;
	END_VAR

	VAR_EXTERNAL
		PLC_TICKS_PER_SEC :	INT;
		PLC_SYS_TICK_CNT :	DINT;
	END_VAR

	VAR
		debug :	BOOL;(*Debug-Mode ON / OFF*)
		N :	INT;(*Debug-Faktor*)
		Offset :	UDINT;(*Debug-Offset*)
		temp :	DWORD := DWORD#1;(*Debug-Offset*)
		mode :	BOOL;(*modus*)
		faktor :	UDINT;(*Systemtakt-Faktor*)
		init :	BOOL;
		v_plc_ticks_per_sec :	UDINT;
		base :	UDINT := UDINT#1000;
	END_VAR

	IF init = FALSE THEN
		v_plc_ticks_per_sec := INT_TO_UDINT(PLC_TICKS_PER_SEC);
		IF v_plc_ticks_per_sec = UDINT#1024 THEN
			faktor := UDINT#1;
			mode := FALSE;
		ELSIF v_plc_ticks_per_sec > UDINT#0 THEN
			IF v_plc_ticks_per_sec <= base THEN
				faktor := base / v_plc_ticks_per_sec;
				mode := FALSE;
			ELSE
				faktor := v_plc_ticks_per_sec / base;
				mode := TRUE;
			END_IF;
		ELSE
			faktor := UDINT#1;
		END_IF;
		init := TRUE;
	END_IF;

	IF mode THEN
		T_PLC_MS := DINT_TO_UDINT(PLC_SYS_TICK_CNT) / faktor;
	ELSE
		T_PLC_MS := DINT_TO_UDINT(PLC_SYS_TICK_CNT) * faktor;
	END_IF;

	IF debug THEN
		T_PLC_MS := (DWORD_TO_UDINT(SHL(UDINT_TO_DWORD(T_PLC_MS),N) OR SHL(temp,N)) - UDINT#1) + Offset;
	END_IF;
END_FUNCTION_BLOCK

FUNCTION _WORD_TO_DINT:DINT
	VAR_INPUT
		IN :	WORD;
	END_VAR
	_WORD_TO_DINT := UINT_TO_DINT(WORD_TO_UINT(IN));
END_FUNCTION

FUNCTION TIME_TO_UDINT2:UDINT
	VAR_INPUT
		X :	TIME;
	END_VAR

	TIME_TO_UDINT2 := DINT_TO_UDINT(TIME_TO_DINT(X));
END_FUNCTION

FUNCTION_BLOCK _RMP_W

	VAR_INPUT
		DIR :	BOOL;
		E :	BOOL := TRUE;
		TR :	TIME;
	END_VAR

	VAR_IN_OUT
		RMP :	WORD;
	END_VAR

	VAR
		T_PLC_MS :	T_PLC_MS_block;
		tx :	UDINT;
		tl :	UDINT;
		ptesss :	DINT;
		init :	BOOL;
		last_dir :	BOOL;
	END_VAR

	T_PLC_MS();
	tx := T_PLC_MS.T_PLC_MS;
	IF E AND init THEN
		(* we need to set tl = tx when direction changes *)
		IF dir XOR last_dir THEN
			tl := tx;
			last_dir := dir;
		END_IF;
		(* check_elapsed time and calculate only if necessary *)
		IF tr > t#0s THEN
			ptesss := DWORD_TO_DINT(UDINT_TO_DWORD(DWORD_TO_UDINT(SHL(UDINT_TO_DWORD(tx-tl), 16)) / TIME_TO_UDINT2(TR)));
		ELSE
			ptesss := DINT#65535;
		END_IF;
		IF ptesss > DINT#0 THEN
			(* perform the ptesss on the ramp *)
			tl := tx;
			(* calculate the ptesss response *)
			IF NOT dir THEN ptesss := - ptesss; END_IF;
			rmp := DINT_TO_WORD(LIMIT(DINT#0, _WORD_TO_DINT(rmp) + ptesss, DINT#65535));
		END_IF;
	ELSE
		tl := tx;
		init := TRUE;
	END_IF;
END_FUNCTION_BLOCK

FUNCTION_BLOCK RMP_W

	VAR_INPUT
		SET :	BOOL;
		PT :	TIME;
		E :	BOOL := TRUE;
		UP :	BOOL := TRUE;
		RST :	BOOL;
	END_VAR

	VAR_OUTPUT
		OUT :	WORD;
		BUSY :	BOOL;
		HIGH :	BOOL;
		LOW :	BOOL;
	END_VAR

	VAR
		rmp :	_RMP_W;
	END_VAR

	rmp(dir := UP, E := E, TR := PT, rmp := out);
	out := rmp.RMP;

	IF RST THEN
		out := WORD#0;
	ELSIF SET THEN
		out := WORD#65535;
	END_IF;

	low := out = WORD#0;
	high := out = WORD#65535;
	busy := NOT (low OR high) AND E;

END_FUNCTION_BLOCK

FUNCTION _WORD_TO_REAL:REAL
	VAR_INPUT
		IN :	WORD;
	END_VAR
	_WORD_TO_REAL := UINT_TO_REAL(WORD_TO_UINT(IN));
END_FUNCTION

FUNCTION_BLOCK FADE
	VAR_INPUT
		IN1 :	REAL;
		IN2 :	REAL;
		F :	BOOL;
		TF :	TIME;
		RST :	BOOL;
	END_VAR

	VAR_OUTPUT
		Y :	REAL;
	END_VAR

	VAR
		rmx :	RMP_W;
	END_VAR
	rmx(rst := rst AND NOT F, set := rst AND F, pt := TF, up := F);
	Y := (in2 - In1) / 65535.0 * _WORD_TO_REAL(rmx.out) + in1;

END_FUNCTION_BLOCK

PROGRAM program0
  VAR

	IN1 :	REAL;
	IN2 :	REAL;
	F   :	BOOL;
	TF  :	TIME;
	RST :	BOOL;

	Y :	REAL;

	func_block : FADE;
  END_VAR
	func_block.IN1 :=IN1;
	func_block.IN2 :=IN2;
	func_block.F   :=F  ;
	func_block.TF  :=TF ;
	func_block.RST :=RST;
	func_block();
	Y := func_block.Y;

END_PROGRAM

CONFIGURATION Config0
	VAR_GLOBAL
		PLC_TICKS_PER_SEC :	INT;
		PLC_SYS_TICK_CNT :	DINT;
	END_VAR
  	RESOURCE Res0 ON PLC
    	TASK task0(INTERVAL := T#20ms,PRIORITY := 0);
    	PROGRAM instance0 WITH task0 : program0;
  	END_RESOURCE
END_CONFIGURATION

(* ---- FF_D2E.ST ---- *)
FUNCTION_BLOCK FF_D2E
	VAR_INPUT
		D0 :	BOOL;
		D1 :	BOOL;
		CLK :	BOOL;
		RST :	BOOL;
	END_VAR

	VAR_OUTPUT
		Q0 :	BOOL;
		Q1 :	BOOL;
	END_VAR

	VAR
		edge :	BOOL;
	END_VAR

	IF rst THEN
		Q0 := FALSE;
		Q1 := FALSE;
	ELSIF clk AND NOT edge THEN
		Q0 := D0;
		Q1 := D1;
	END_IF;
	edge := CLK;

END_FUNCTION_BLOCK

PROGRAM program0
  VAR
	D0  :	BOOL;
	D1  :	BOOL;
	CLK :	BOOL;
	RST :	BOOL;

	Q0 :	BOOL;
	Q1 :	BOOL;

	func_block : FF_D2E;
  END_VAR
	func_block.D0  :=D0 ;
	func_block.D1  :=D1 ;
	func_block.CLK :=CLK;
	func_block.RST :=RST;
	func_block();
	Q0 := func_block.Q0;
	Q1 := func_block.Q1;
END_PROGRAM

CONFIGURATION Config0
  RESOURCE Res0 ON PLC
    TASK task0(INTERVAL := T#20ms,PRIORITY := 0);
    PROGRAM instance0 WITH task0 : program0;
  END_RESOURCE
END_CONFIGURATION

(* ---- FF_D4E.ST ---- *)
FUNCTION_BLOCK FF_D4E
	VAR_INPUT
		D0 :	BOOL;
		D1 :	BOOL;
		D2 :	BOOL;
		D3 :	BOOL;
		CLK :	BOOL;
		RST :	BOOL;
	END_VAR

	VAR_OUTPUT
		Q0 :	BOOL;
		Q1 :	BOOL;
		Q2 :	BOOL;
		Q3 :	BOOL;
	END_VAR

	VAR
		edge :	BOOL;
	END_VAR

	IF rst THEN
		Q0 := FALSE;
		Q1 := FALSE;
		Q2 := FALSE;
		Q3 := FALSE;
	ELSIF clk AND NOT edge THEN
		Q0 := D0;
		Q1 := D1;
		Q2 := D2;
		Q3 := D3;
	END_IF;
	edge := CLK;
END_FUNCTION_BLOCK

PROGRAM program0
  VAR
		D0  :	BOOL;
		D1  :	BOOL;
		D2  :	BOOL;
		D3  :	BOOL;
		CLK :	BOOL;
		RST :	BOOL;

		Q0 :	BOOL;
		Q1 :	BOOL;
		Q2 :	BOOL;
		Q3 :	BOOL;

	func_block : FF_D4E;
  END_VAR
	func_block.D0 :=D0 ;
	func_block.D1 :=D1 ;
	func_block.D2 :=D2 ;
	func_block.D3 :=D3 ;
	func_block.CLK:=CLK;
	func_block.RST:=RST;
	func_block();
	Q0 := func_block.Q0;
	Q1 := func_block.Q1;
	Q2 := func_block.Q2;
	Q3 := func_block.Q3;
END_PROGRAM

CONFIGURATION Config0
  RESOURCE Res0 ON PLC
    TASK task0(INTERVAL := T#20ms,PRIORITY := 0);
    PROGRAM instance0 WITH task0 : program0;
  END_RESOURCE
END_CONFIGURATION

(* ---- FF_DRE.ST ---- *)
FUNCTION_BLOCK FF_DRE
	VAR_INPUT
		SET :	BOOL;
		D :	BOOL;
		CLK :	BOOL;
		RST :	BOOL;
	END_VAR

	VAR_OUTPUT
		Q :	BOOL;
	END_VAR

	VAR
		edge :	BOOL;
	END_VAR

	IF rst OR set THEN
		Q := NOT rst;
	ELSIF clk AND NOT edge THEN
		Q := D;
	END_IF;
	edge := CLK;

END_FUNCTION_BLOCK

PROGRAM program0
  VAR
	SET :	BOOL;
	D   :	BOOL;
	CLK :	BOOL;
	RST :	BOOL;

	Q :	BOOL;

	func_block : FF_DRE;
  END_VAR
	func_block.SET:=SET;
	func_block.D  :=D  ;
	func_block.CLK:=CLK;
	func_block.RST:=RST;
	func_block();
	Q:= func_block.Q;
END_PROGRAM

CONFIGURATION Config0
  RESOURCE Res0 ON PLC
    TASK task0(INTERVAL := T#20ms,PRIORITY := 0);
    PROGRAM instance0 WITH task0 : program0;
  END_RESOURCE
END_CONFIGURATION

(* ---- FF_JKE.ST ---- *)
FUNCTION_BLOCK FF_JKE
	VAR_INPUT
		SET :	BOOL;
		J :	BOOL;
		CLK :	BOOL;
		K :	BOOL;
		RST :	BOOL;
	END_VAR

	VAR_OUTPUT
		Q :	BOOL;
	END_VAR

	VAR
		edge :	BOOL;
	END_VAR

	IF rst OR set THEN
		Q := NOT rst;
	ELSIF clk AND NOT edge THEN
		IF J XOR K THEN Q := J;
		ELSE Q := K XOR Q;
		END_IF;
	END_IF;
	edge := CLK;

END_FUNCTION_BLOCK

PROGRAM program0
  VAR
		SET :	BOOL;
		J   :	BOOL;
		CLK :	BOOL;
		K   :	BOOL;
		RST :	BOOL;

		Q :	BOOL;

	func_block : FF_JKE;
  END_VAR
	func_block.SET :=SET;
	func_block.J   :=J  ;
	func_block.CLK :=CLK;
	func_block.K   :=K  ;
	func_block.RST :=RST;
	func_block();
	Q := func_block.Q;
END_PROGRAM

CONFIGURATION Config0
  RESOURCE Res0 ON PLC
    TASK task0(INTERVAL := T#20ms,PRIORITY := 0);
    PROGRAM instance0 WITH task0 : program0;
  END_RESOURCE
END_CONFIGURATION

(* ---- FF_RSE.ST ---- *)
FUNCTION_BLOCK FF_RSE
	VAR_INPUT
		CS :	BOOL;
		CR :	BOOL;
		RST :	BOOL;
	END_VAR

	VAR_OUTPUT
		Q :	BOOL;
	END_VAR

	VAR
		es :	BOOL;
		er :	BOOL;
	END_VAR

	IF rst THEN
		(* asynchronous reset *)
		Q := FALSE;
	ELSIF CR AND NOT er THEN
		(* rising edge on CR *)
		Q := FALSE;
	ELSIF CS AND NOT es THEN
		(* rising edge on CS *)
		Q := TRUE;
	END_IF;

	es := CS;
	er := CR;
END_FUNCTION_BLOCK

PROGRAM program0
  VAR
	CS  :	BOOL;
	CR  :	BOOL;
	RST :	BOOL;

	Q :	BOOL;

	func_block : FF_RSE;
  END_VAR
	func_block.CS  :=CS ;
	func_block.CR  :=CR ;
	func_block.RST :=RST;
	func_block();
	Q := func_block.Q;
END_PROGRAM

CONFIGURATION Config0
  RESOURCE Res0 ON PLC
    TASK task0(INTERVAL := T#20ms,PRIORITY := 0);
    PROGRAM instance0 WITH task0 : program0;
  END_RESOURCE
END_CONFIGURATION

(* ---- FIFO_16.ST ---- *)
TYPE
	oscat_ardw_0_15             : ARRAY [0..15]   OF DWORD;
END_TYPE

FUNCTION INC1:INT

	VAR_INPUT
		X :	INT;
		N :	INT;
	END_VAR

	IF X >= N - 1 THEN
		INC1 := 0;
	ELSE
		INC1 := X + 1;
	END_IF;
END_FUNCTION

FUNCTION_BLOCK FIFO_16
	VAR_INPUT
		DIN :	DWORD;
		E :	BOOL := TRUE;
		RD :	BOOL;
		WD :	BOOL;
		RST :	BOOL;
	END_VAR

	VAR_OUTPUT
		DOUT :	DWORD;
		EMPTY :	BOOL := TRUE;
		FULL :	BOOL;
	END_VAR

	VAR
		fifo :	oscat_ardw_0_15;
		pr :	INT;
		pw :	INT;
	END_VAR

	IF RST THEN
		pw := pr;
		FULL := FALSE;
		EMPTY := TRUE;
		Dout := DWORD#0;
	ELSIF E THEN
		IF NOT EMPTY AND RD THEN
			Dout := fifo[pr];
			pr := INC1(pr,16);
			EMPTY := pr = pw;
			FULL := FALSE;
		END_IF;
		IF NOT FULL AND WD THEN
			fifo[pw] := Din;
			pw := INC1(pw,16);
			FULL := pw = pr;
			EMPTY := FALSE;
		END_IF;
	END_IF;
END_FUNCTION_BLOCK

PROGRAM program0
  VAR
	DIN :	DWORD;
	E   :	BOOL;
	RD  :	BOOL;
	WD  :	BOOL;
	RST :	BOOL;

	DOUT  :	DWORD;
	EMPTY :	BOOL;
	FULL  :	BOOL;

	func_block : FIFO_16;
  END_VAR
	func_block.DIN :=DIN;
	func_block.E   :=E  ;
	func_block.RD  :=RD ;
	func_block.WD  :=WD ;
	func_block.RST :=RST;
	func_block();
	DOUT := func_block.DOUT ;
	EMPTY:= func_block.EMPTY;
	FULL := func_block.FULL ;
END_PROGRAM

CONFIGURATION Config0
  RESOURCE Res0 ON PLC
    TASK task0(INTERVAL := T#20ms,PRIORITY := 0);
    PROGRAM instance0 WITH task0 : program0;
  END_RESOURCE
END_CONFIGURATION

(* ---- FIFO_32.ST ---- *)
TYPE
	oscat_ardw_0_31             : ARRAY [0..31]   OF DWORD;
END_TYPE

FUNCTION INC1:INT

	VAR_INPUT
		X :	INT;
		N :	INT;
	END_VAR

	IF X >= N - 1 THEN
		INC1 := 0;
	ELSE
		INC1 := X + 1;
	END_IF;
END_FUNCTION

FUNCTION_BLOCK FIFO_32

	VAR_INPUT
		DIN :	DWORD;
		E :	BOOL := TRUE;
		RD :	BOOL;
		WD :	BOOL;
		RST :	BOOL;
	END_VAR

	VAR_OUTPUT
		DOUT :	DWORD;
		EMPTY :	BOOL := TRUE;
		FULL :	BOOL;
	END_VAR

	VAR
		fifo :	oscat_ardw_0_31;
		pr :	INT;
		pw :	INT;
	END_VAR

	IF RST THEN
		pw := pr;
		FULL := FALSE;
		EMPTY := TRUE;
		Dout := DWORD#0;
	ELSIF E THEN
		IF NOT EMPTY AND RD THEN
			Dout := fifo[pr];
			pr := INC1(pr,32);
			EMPTY := pr = pw;
			FULL := FALSE;
		END_IF;
		IF NOT FULL AND WD THEN
			fifo[pw] := Din;
			pw := INC1(pw,32);
			FULL := pw = pr;
			EMPTY := FALSE;
		END_IF;
	END_IF;

END_FUNCTION_BLOCK

PROGRAM program0
  VAR
	DIN :	DWORD;
	E   :	BOOL;
	RD  :	BOOL;
	WD  :	BOOL;
	RST :	BOOL;

	DOUT  :	DWORD;
	EMPTY :	BOOL;
	FULL  :	BOOL;

	func_block : FIFO_32;
  END_VAR
	func_block.DIN :=DIN;
	func_block.E   :=E  ;
	func_block.RD  :=RD ;
	func_block.WD  :=WD ;
	func_block.RST :=RST;
	func_block();
	DOUT := func_block.DOUT ;
	EMPTY:= func_block.EMPTY;
	FULL := func_block.FULL ;
END_PROGRAM

CONFIGURATION Config0
  RESOURCE Res0 ON PLC
    TASK task0(INTERVAL := T#20ms,PRIORITY := 0);
    PROGRAM instance0 WITH task0 : program0;
  END_RESOURCE
END_CONFIGURATION

(* ---- FILE_BLOCK.ST ---- *)
TYPE
  oscat_FILE_SERVER_DATA : STRUCT
	FILE_OPEN	: BOOL;
    FILENAME 	: STRING;
    MODE	 	: BYTE;
    OFFSET   	: UDINT;
    FILE_SIZE   : UDINT;
    AUTO_CLOSE	: TIME;
    ERROR	 	: BYTE;
  END_STRUCT;

  oscat_NW_BUF_LONG  : ARRAY [0..4095] OF BYTE;
  oscat_NETWORK_BUFFER :
  STRUCT
    SIZE   : UINT;
    BUFFER : oscat_NW_BUF_LONG;
  END_STRUCT;
END_TYPE

FUNCTION_BLOCK FILE_BLOCK

	VAR_IN_OUT
		MODE :	BYTE;
		FILENAME :	STRING;
		FSD :	oscat_FILE_SERVER_DATA;
		PT :	oscat_NETWORK_BUFFER;
	END_VAR

	VAR_INPUT
		POS :	UDINT;
	END_VAR

	VAR_OUTPUT
		ERROR :	BYTE;
		DATA :	BYTE;
	END_VAR

	VAR
		stepp :	INT;
		i :	INT;
		data_start :	UDINT;
		data_stop :	UDINT;
	END_VAR

	CASE stepp OF
	0:	IF MODE > BYTE#0 THEN
			ERROR := BYTE#0;
			IF FSD.FILE_OPEN AND (FSD.FILE_SIZE = UDINT#0 OR POS >= FSD.FILE_SIZE) THEN
				ERROR := BYTE#255;
				MODE := BYTE#0;
			ELSIF POS < data_start OR POS > data_stop OR NOT FSD.FILE_OPEN THEN
				FSD.FILENAME := FILENAME;
				FSD.MODE := BYTE#1;
				FSD.OFFSET := POS;
				PT.SIZE := UINT#65535;
				data_start := UDINT#0;
				data_stop := UDINT#0;
				stepp := 10;
			ELSE
				i := UDINT_TO_INT(POS - data_start);
				DATA := PT.BUFFER[i];
				MODE := BYTE#0;
			END_IF;
		END_IF;

	10:	IF FSD.MODE = BYTE#0 THEN
			IF FSD.ERROR > BYTE#0 THEN
				ERROR := FSD.ERROR;
				MODE := BYTE#0;
			ELSE
				data_start := POS;
				data_stop := POS + UINT_TO_UDINT(PT.SIZE) - UDINT#1;
			END_IF;
			stepp := 0;
		END_IF;
	END_CASE;
END_FUNCTION_BLOCK

PROGRAM program0
	VAR
		MODE :	BYTE;
		FILENAME :	STRING;
		FSD :	oscat_FILE_SERVER_DATA;
		PT :	oscat_NETWORK_BUFFER;
		POS :	UDINT;
		ERROR :	BYTE;
		DATA :	BYTE;

		func_block : FILE_BLOCK;
	END_VAR
	func_block.MODE    :=MODE    ;
	func_block.FILENAME:=FILENAME;
	func_block.FSD     :=FSD     ;
	func_block.PT      :=PT      ;
	func_block.POS     :=POS     ;
	func_block();
	MODE    := func_block.MODE    ;
	FILENAME:= func_block.FILENAME;
	FSD     := func_block.FSD     ;
	PT      := func_block.PT      ;
	ERROR   := func_block.ERROR;
	DATA    := func_block.DATA;

END_PROGRAM

CONFIGURATION Config0
  RESOURCE Res0 ON PLC
    TASK task0(INTERVAL := T#20ms,PRIORITY := 0);
    PROGRAM instance0 WITH task0 : program0;
  END_RESOURCE
END_CONFIGURATION

(* ---- FILE_PATH_SPLIT.ST ---- *)
TYPE
  oscat_STRING250             : STRING;
  oscat_STRING1             : STRING;
  oscat_STRING80             : STRING;
  oscat_STRING3             : STRING;
  oscat_NW_BUF_LONG  : ARRAY [0..4095] OF BYTE;
  PRINTF_DATA_250  	:  ARRAY [1..11]  OF oscat_STRING250;
  PRINTF_DATA_80 	:  ARRAY [1..11]  OF oscat_STRING80;
  LOG_250       	:  ARRAY [0..400] OF oscat_STRING250;
  LOG_80    		:  ARRAY [0..400] OF oscat_STRING80;
  LOG_OPTION		:  ARRAY [0..400] OF DWORD;

  us_LOG_CONTROL :
  STRUCT
    NEW_MSG              : oscat_STRING250;    (*W neue Nachricht f�r den Datenbuffer   *)
	NEW_MSG_OPTION 		 : DWORD;
    LEVEL                : BYTE;
	SIZE                 : INT;                (*R Anzahl der Strings im LOG_DATA       *)
	RESET                : BOOL;               (*W Nachrichtenbuffer l�schen            *)
    PRINTF               : PRINTF_DATA_250;    (*W Array PRINTF Parameter               *)
    MSG                  : LOG_250;            (*I Array Message                        *)
    MSG_OPTION           : LOG_OPTION;     	   (*I Array Message Option                 *)
	UPDATE_COUNT         : UINT;               (*R Updatez�hler                         *)
    IDX                  : INT;                (*R aktueller Nachrichten-Index          *)
	RING_MODE            : BOOL;               (*I Buffer�berlauf erkannt               *)
  END_STRUCT;

  us_LOG_CONTROL_80 :
  STRUCT
    NEW_MSG              : oscat_STRING80;     (*W neue Nachricht f�r den Datenbuffer   *)
	NEW_MSG_OPTION 		 : DWORD;
    LEVEL                : BYTE;
	SIZE                 : INT;                (*R Anzahl der Strings im LOG_DATA       *)
	RESET                : BOOL;               (*W Nachrichtenbuffer l�schen            *)
    PRINTF               : PRINTF_DATA_80;     (*W Array PRINTF Parameter               *)
    MSG                  : LOG_80;             (*I Array Message                        *)
    MSG_OPTION           : LOG_OPTION;     	   (*I Array Message Option                 *)
	UPDATE_COUNT         : UINT;               (*R Updatez�hler                         *)
    IDX                  : INT;                (*R aktueller Nachrichten-Index          *)
	RING_MODE            : BOOL;               (*I Buffer�berlauf erkannt               *)
  END_STRUCT;

  LINE_ARRAY 			: ARRAY [1..40] OF INT;

  us_LOG_VIEWPORT :
    STRUCT
     LINE_ARRAY          : LINE_ARRAY;
     COUNT               : INT;                (* Anzahl der sichtbaren Nachtrichten   *)
	 UPDATE_COUNT        : UINT;               (* Updatez�hler                         *)
     MOVE_TO_X           : INT;                (* Steuerung der Nachrichtenanzeige     *)
     UPDATE              : BOOL;               (* Daten wurden ge�ndert -> neuzeichnen *)
  END_STRUCT;

  oscat_FILE_SERVER_DATA : STRUCT
	FILE_OPEN	: BOOL;
    FILENAME 	: STRING;
    MODE	 	: BYTE;
    OFFSET   	: UDINT;
    FILE_SIZE   : UDINT;
    AUTO_CLOSE	: TIME;
    ERROR	 	: BYTE;
  END_STRUCT;

  oscat_FILE_PATH_DATA : STRUCT
	DRIVE : oscat_string3;
	DIRECTORY : oscat_string250;
	FILENAME : STRING;
  END_STRUCT;

  oscat_UNI_CIRCULAR_BUFFER_DATA : STRUCT
	D_MODE : INT;
	D_HEAD : WORD;
	D_STRING : oscat_string250;
	D_REAL : REAL;
	D_DWORD : DWORD;
	BUF_SIZE : INT;
	BUF_COUNT : INT;
	BUF_USED : USINT;
	BUF : oscat_NW_BUF_LONG;
	_GetStart : INT;
	_GetEnd : INT;
	_Last : INT;
	_First : INT;
  END_STRUCT;

  oscat_DLOG_DATA : STRUCT
	STORE_TYPE : BYTE;
	ADD_HEADER : BOOL;
	ADD_DATA : BOOL;
	ADD_DATA_REQ : BOOL;
	CLOCK_TRIG : BOOL;
	ID_MAX : USINT;
	DTI : UDINT;
	UCB : oscat_UNI_CIRCULAR_BUFFER_DATA;
	NEW_FILE : STRING;
	NEW_FILE_RTRIG : BOOL;
  END_STRUCT;

END_TYPE

FUNCTION_BLOCK FILE_PATH_SPLIT_Block

	VAR_INPUT
		FILENAME :	oscat_STRING250;
	END_VAR

	VAR_OUTPUT
		FILE_PATH_SPLIT :	BOOL;
	END_VAR

	VAR_IN_OUT
		X :	oscat_FILE_PATH_DATA;
	END_VAR

	VAR
		b :	INT;
		c :	INT;
		d :	oscat_STRING1;
		p1 :	INT;
		p2 :	INT;
	END_VAR

	X.DRIVE := '';
	X.DIRECTORY := '';
	X.FILENAME := '';
	p1 := 0;
	p2 := 0;
	c := LEN(FILENAME);
	IF c = 0 THEN
		FILE_PATH_SPLIT := FALSE;
		RETURN;
	END_IF;

	FOR b := 1 TO c DO
		d := MID(FILENAME, 1, b);
		IF EQ_STRING(d,':') THEN
			p1 := b;
		ELSIF EQ_STRING(d,'/') OR EQ_STRING(d,'\') THEN
			p2 := b;
		END_IF;
	END_FOR;

	IF p1 = 2 THEN
		X.DRIVE := LEFT(FILENAME,p1);
	END_IF;

	IF p2 > 0 AND p2 > p1 THEN
		X.DIRECTORY := MID(FILENAME,p2-p1,p1+1);
	END_IF;

	X.FILENAME := RIGHT(FILENAME,c - MAX (p1,p2));
	FILE_PATH_SPLIT := TRUE;

END_FUNCTION_BLOCK

PROGRAM program0
	VAR
		FILENAME :	oscat_STRING250;
		FILE_PATH_SPLIT :	BOOL;
		X :	oscat_FILE_PATH_DATA;

		func_block : FILE_PATH_SPLIT_Block;
	END_VAR
	func_block.FILENAME := FILENAME;
	func_block.X := X;

	func_block();
	FILE_PATH_SPLIT  := func_block.FILE_PATH_SPLIT;
	X  := func_block.X;
END_PROGRAM

CONFIGURATION Config0
	RESOURCE Res0 ON PLC
		TASK task0(INTERVAL := T#20ms,PRIORITY := 0);
		PROGRAM instance0 WITH task0 : program0;
	END_RESOURCE
END_CONFIGURATION

(* ---- FILE_SERVER.ST ---- *)
FUNCTION_BLOCK FILE_SERVER_Block

	VAR
		buf_size :	UDINT := UDINT#4096;
		handle :	UINT;
		read_max_length :	UDINT;
		file_position :	UDINT;
		used_filename :	STRING;
		close_time :	TIME;
		length_read :	UDINT;
		write_length :	UDINT;
		length_written :	UDINT;
		open_handle :	UINT;
		seek_mode :	UINT;
		seek_position :	UDINT;
		tell_position :	UDINT;
	END_VAR

	VAR
		last_mode :	BYTE;
		command :	BYTE;
		error_code :	BYTE;
		error :	BOOL;
		file_change :	BOOL;
		step :	INT;
		t_diff :	TIME;
		tx_last :	TIME;
		tx :	TIME;
	END_VAR

	VAR_IN_OUT
		FSD :	oscat_FILE_SERVER_DATA;
		PT :	oscat_NETWORK_BUFFER;
	END_VAR

	VAR
		FILE_REMOVE :	FILE_REMOVE;
		FILE_OPEN :	FILE_OPEN;
		FILE_SEEK :	FILE_SEEK;
		FILE_TELL :	FILE_TELL;
		FILE_CLOSE :	FILE_CLOSE;
		FILE_READ :	FILE_READ;
		FILE_WRITE :	FILE_WRITE;
		T_PLC_MS :	T_PLC_MS;
	END_VAR

	T_PLC_MS();
	tx := UDINT_TO_TIME(T_PLC_MS.T_PLC_MS);
	t_diff := tx - tx_last;
	tx_last := tx;

	CASE step OF
	0:
		IF FSD.MODE = LIMIT(BYTE#1,FSD.MODE,BYTE#5) THEN
			close_time := T#1ms;
			IF handle = UINT#00 AND FSD.MODE <= BYTE#3 THEN
				step := 100;
			ELSE
				IF EQ_STRING(used_filename, FSD.FILENAME) AND FSD.MODE = last_mode THEN
					step := 200;
				ELSE
					step := 32000;
					file_change := FSD.MODE <> BYTE#5;
				END_IF;
			END_IF;
		ELSIF handle > UINT#0 THEN
			IF FSD.AUTO_CLOSE > T#0s THEN
				close_time := close_time + t_diff;
				IF close_time > FSD.AUTO_CLOSE THEN
					step := 32000;
				END_IF;
			END_IF;
		END_IF;

	100:
		IF FSD.MODE = BYTE#3 OR FSD.MODE = BYTE#4 THEN
			command := BYTE#7;
			step := 110;
		ELSE
			step := 120;
		END_IF;

	110:
		IF command = BYTE#0  THEN
			IF (FSD.MODE = BYTE#4) OR (error and error_code <> BYTE#143) THEN
				step := 30000;
			ELSE
				step := 120;
			END_IF;
		END_IF;

	120:
		command := BYTE#1;
		last_mode := FSD.MODE;
		step := 122;

	122:
		IF command = BYTE#0 THEN
			IF error THEN
				step := 30000;
			ELSE

				close_time := T#1ms;
				handle := open_handle;
				used_filename := FSD.FILENAME;
				file_position := UDINT#4294967295;
				FSD.FILE_SIZE := UDINT#0;
				step := 125;
			END_IF;
		END_IF;

	125:
		seek_mode := UINT#2;
		seek_position := UDINT#0;
		command := BYTE#5;
		step := 130;

	130:
		IF command = BYTE#0 THEN
			IF Error THEN
				step := 30000;
			ELSE
				step := 140;
			END_IF;
		END_IF;

	140:
		command := BYTE#6;
		step := 150;

	150:
		IF command = BYTE#0 THEN
			IF Error THEN
				step := 30000;
			ELSE
				FSD.FILE_SIZE := tell_position;
				file_position := tell_position;
				FSD.FILE_OPEN := TRUE;
				step := 200;
			END_IF;
		END_IF;

	200:
		IF FSD.OFFSET > FSD.FILE_SIZE THEN
			error_code := BYTE#255;
			step := 30000;
		ELSIF FSD.OFFSET <> file_position THEN
			command := BYTE#5;
			seek_mode := UINT#0;
			seek_position := FSD.OFFSET;
			step := 210;
		ELSE
			step := 300;
		END_IF;

	210:
		IF command = BYTE#0 THEN
			file_position := seek_position;
			IF Error THEN
				step := 30000;
			ELSE
				step := 300;
			END_IF;
		END_IF;

	300:
		IF FSD.MODE = BYTE#1 THEN
			step := 400;
		ELSE
			step := 500;
		END_IF;

	400:
		IF UINT_TO_UDINT(PT.SIZE) > buf_size THEN
			read_max_length := buf_size;
		ELSE
			read_max_length := UINT_TO_UDINT(PT.SIZE);
		END_IF;

		IF file_position + read_max_length > FSD.FILE_SIZE THEN
			read_max_length := FSD.FILE_SIZE - file_position;
		END_IF;

		IF read_max_length > UDINT#0 THEN
			command := BYTE#3;
			step := INT#410;
		ELSE
			PT.SIZE := UINT#0;
			step := 30000;
		END_IF;

	410:
		IF command = BYTE#0 THEN
			PT.SIZE := UDINT_TO_UINT(length_read);
			IF NOT Error THEN
				file_position := file_position + length_read;
				FSD.OFFSET := file_position;
			END_IF;
			step := 30000;
		END_IF;

	500:
		IF UINT_TO_UDINT(PT.SIZE) > buf_size THEN
			write_length := buf_size;
		ELSE
			write_length := UINT_TO_UDINT(PT.SIZE);
		END_IF;

		IF write_length > UDINT#0 THEN
			command := BYTE#4;
			step := INT#510;
		ELSE
			step := 30000;
		END_IF;

	510:
		IF command = BYTE#0 THEN
			IF NOT Error THEN
				file_position := file_position + length_written;
				FSD.OFFSET := file_position;
				IF file_position > FSD.FILE_SIZE THEN
					FSD.FILE_SIZE := file_position;
				END_IF;
			END_IF;
			step := 30000;
		END_IF;

	30000:
		FSD.MODE := BYTE#0;
		FSD.ERROR := error_code;
		step := 0;

	32000:
		close_time := T#0s;
		IF handle > UINT#0 THEN
			command := BYTE#2;
		END_IF;
		step := 32100;

	32100:
		IF command = BYTE#0 THEN
			FSD.FILE_OPEN := FALSE;
			file_position := UDINT#0;
			FSD.FILE_SIZE := UDINT#0;
			FSD.OFFSET := UDINT#0;
			used_filename := '';
			handle := UINT#00;

			IF file_change THEN
				file_change := FALSE;
				step := 100;
			ELSE
				step := 30000;
			END_IF;
		END_IF;

	END_CASE;

	FILE_OPEN.Execute := command = BYTE#1;
	FILE_OPEN.Name := FSD.FILENAME;
	FILE_OPEN();
	open_handle := FILE_OPEN.Handle;

	IF command = BYTE#1 THEN
		IF FILE_OPEN.Done THEN
			error := FILE_OPEN.Error;
			command := BYTE#0;
			error_code := SEL_BYTE(error,BYTE#00,UINT_TO_BYTE(FILE_OPEN.ErrorID));
		END_IF;
	END_IF;

	FILE_CLOSE.Execute := command = BYTE#2;
	FILE_CLOSE.Handle := Handle;
	FILE_CLOSE();

	IF command = BYTE#2 THEN
		IF FILE_CLOSE.Done THEN
			error := FILE_CLOSE.Error;
			command := BYTE#0;
			error_code := SEL_BYTE(error,BYTE#00,UINT_TO_BYTE(FILE_CLOSE.ErrorID + UINT#10));
		END_IF;
	END_IF;

	FILE_READ.Execute := command = BYTE#3;
	FILE_READ.Handle := handle;
	FILE_READ.MaxLength := read_max_length;
	FILE_READ.Buffer := PT.BUFFER;
	FILE_READ();
	PT.BUFFER := FILE_READ.Buffer;

	IF command = BYTE#3 THEN
		IF FILE_READ.Done THEN
			error := FILE_READ.Error;
			command := BYTE#0;
			length_read :=  FILE_READ.LengthRead;
			error_code := SEL_BYTE(error,BYTE#00,UINT_TO_BYTE(FILE_READ.ErrorID + UINT#40));
		END_IF;
	END_IF;

	FILE_WRITE.Execute   := command = BYTE#4;
	FILE_WRITE.Handle    := handle;
	FILE_WRITE.Length    := write_length ;
	FILE_WRITE.Buffer    := PT.BUFFER;
	FILE_WRITE();
	PT.BUFFER := FILE_WRITE.Buffer;

	IF command = BYTE#4 THEN
		IF FILE_WRITE.Done THEN
			error := FILE_WRITE.Error;
			command := BYTE#0;
			length_written := write_length;
			error_code := SEL_BYTE(error,BYTE#00,UINT_TO_BYTE(FILE_WRITE.ErrorID + UINT#70));
		END_IF;
	END_IF;

	FILE_SEEK.Execute  := command = BYTE#5;
	FILE_SEEK.Handle   := handle;
	FILE_SEEK.Mode     := seek_mode;
	FILE_SEEK.Position := UDINT_TO_DINT(seek_position);
	FILE_SEEK();

	IF command = BYTE#5 THEN
		IF FILE_SEEK.Done THEN
			error := FILE_SEEK.Error;
			command := BYTE#0;
			error_code := SEL_BYTE(error,BYTE#00,UINT_TO_BYTE(FILE_SEEK.ErrorID + UINT#100));
		END_IF;
	END_IF;

	FILE_TELL.Execute := command = BYTE#6;
	FILE_TELL.Handle := handle;
	FILE_TELL();

	IF command = BYTE#6 THEN
		IF FILE_TELL.Done THEN
			error := FILE_TELL.Error;
			command := BYTE#0;
			tell_position := DINT_TO_UDINT(FILE_TELL.Position);
			error_code := SEL_BYTE(error,BYTE#00,UINT_TO_BYTE(FILE_TELL.ErrorID + UINT#130));
		END_IF;
	END_IF;

	FILE_REMOVE.Execute := command = BYTE#7;
	FILE_REMOVE.Name := FSD.FILENAME;
	FILE_REMOVE();

	IF command = BYTE#7 THEN
		IF FILE_REMOVE.Done THEN
			error := FILE_REMOVE.Error;
			command := BYTE#0;
			error_code := SEL_BYTE(error,BYTE#00,UINT_TO_BYTE(FILE_REMOVE.ErrorID + UINT#140));
		END_IF;
	END_IF;

END_FUNCTION_BLOCK

PROGRAM program0
	VAR
		FSD :	oscat_FILE_SERVER_DATA;
		PT :	oscat_NETWORK_BUFFER;

		func_block : FILE_SERVER_Block;
	END_VAR
	func_block.FSD := FSD;
	func_block.PT := PT;

	func_block();
	FSD  := func_block.FSD;
	PT  := func_block.PT;
END_PROGRAM

CONFIGURATION Config0
	RESOURCE Res0 ON PLC
		TASK task0(INTERVAL := T#20ms,PRIORITY := 0);
		PROGRAM instance0 WITH task0 : program0;
	END_RESOURCE
END_CONFIGURATION

(* ---- FILL.ST ---- *)
FUNCTION_BLOCK CHR_TO_STRING_Block
	VAR_INPUT
		C :	BYTE;
	END_VAR

	VAR_OUTPUT
		CHR_TO_STRING :	STRING;
	END_VAR

	CHR_TO_STRING := BYTE_TO_STRING(C);

END_FUNCTION_BLOCK

FUNCTION BIT_OF_DWORD : BOOL
  VAR_INPUT
    IN : DWORD;
    N : INT;
  END_VAR

  BIT_OF_DWORD := (SHR(in,N) AND 16#00000001) > 0;
  (* from OSCAT library; www.oscat.de  *)
END_FUNCTION

FUNCTION_BLOCK FILL_Block
	VAR_INPUT
		C :	BYTE;
		L :	INT;
	END_VAR

	VAR_OUTPUT
		FILL :	STRING;
	END_VAR

	VAR
		N :	BYTE;
		I :	INT;
		sx :	STRING;
		CHR_TO_STRING :	CHR_TO_STRING_Block;
		FILL_tmp :	STRING;
	END_VAR

	CHR_TO_STRING(C:=c);
	Sx:=CHR_TO_STRING.CHR_TO_STRING;
	(* create string *)
	N := INT_TO_BYTE(LIMIT(0,L,80));
	(* create a string of characters to be connected to str *)
	FILL := '';
	FOR i := 1 TO 8 DO
		FILL_tmp := FILL;
		FILL := CONCAT(FILL_tmp,FILL);
		IF BIT_OF_DWORD(BYTE_TO_DWORD(N),7) THEN FILL := CONCAT(FILL,Sx); END_IF;
		N := SHL(N,1);
	END_FOR;
END_FUNCTION_BLOCK

PROGRAM program0
  VAR
	C :	BYTE;
	L :	INT;

	FILL :	STRING;

	func_block : FILL_Block;
  END_VAR
	func_block.C  :=C ;
	func_block.L  :=L ;
	func_block();
	FILL := func_block.FILL;
END_PROGRAM

CONFIGURATION Config0
  RESOURCE Res0 ON PLC
    TASK task0(INTERVAL := T#20ms,PRIORITY := 0);
    PROGRAM instance0 WITH task0 : program0;
  END_RESOURCE
END_CONFIGURATION

(* ---- FILTER_DW.ST ---- *)
FUNCTION_BLOCK T_PLC_MS_block
	VAR_OUTPUT
		T_PLC_MS :	UDINT;
	END_VAR

	VAR_EXTERNAL
		PLC_TICKS_PER_SEC :	INT;
		PLC_SYS_TICK_CNT :	DINT;
	END_VAR

	VAR
		debug :	BOOL;(*Debug-Mode ON / OFF*)
		N :	INT;(*Debug-Faktor*)
		Offset :	UDINT;(*Debug-Offset*)
		temp :	DWORD := DWORD#1;(*Debug-Offset*)
		mode :	BOOL;(*modus*)
		faktor :	UDINT;(*Systemtakt-Faktor*)
		init :	BOOL;
		v_plc_ticks_per_sec :	UDINT;
		base :	UDINT := UDINT#1000;
	END_VAR

	IF init = FALSE THEN
		v_plc_ticks_per_sec := INT_TO_UDINT(PLC_TICKS_PER_SEC);
		IF v_plc_ticks_per_sec = UDINT#1024 THEN
			faktor := UDINT#1;
			mode := FALSE;
		ELSIF v_plc_ticks_per_sec > UDINT#0 THEN
			IF v_plc_ticks_per_sec <= base THEN
				faktor := base / v_plc_ticks_per_sec;
				mode := FALSE;
			ELSE
				faktor := v_plc_ticks_per_sec / base;
				mode := TRUE;
			END_IF;
		ELSE
			faktor := UDINT#1;
		END_IF;
		init := TRUE;
	END_IF;

	IF mode THEN
		T_PLC_MS := DINT_TO_UDINT(PLC_SYS_TICK_CNT) / faktor;
	ELSE
		T_PLC_MS := DINT_TO_UDINT(PLC_SYS_TICK_CNT) * faktor;
	END_IF;

	IF debug THEN
		T_PLC_MS := (DWORD_TO_UDINT(SHL(UDINT_TO_DWORD(T_PLC_MS),N) OR SHL(temp,N)) - UDINT#1) + Offset;
	END_IF;

END_FUNCTION_BLOCK

FUNCTION _DWORD_TO_REAL:REAL
	VAR_INPUT
		IN :	DWORD;
	END_VAR

	_DWORD_TO_REAL := UDINT_TO_REAL(DWORD_TO_UDINT(IN));
END_FUNCTION

FUNCTION _REAL_TO_DWORD: DWORD

  VAR_INPUT
    X :	REAL;
  END_VAR

  IF REAL_TO_DWORD(0.5) = DWORD#1 THEN
    _REAL_TO_DWORD := REAL_TO_DWORD(x);
  ELSIF X > 0.0 THEN
    _REAL_TO_DWORD := REAL_TO_DWORD(x+0.5);
  ELSIF X < 0.0 THEN
    _REAL_TO_DWORD := REAL_TO_DWORD(x-0.5);
  ELSE
    _REAL_TO_DWORD := DWORD#0;
  END_IF;
END_FUNCTION

FUNCTION_BLOCK FILTER_DW

	VAR_INPUT
		X :	DWORD;
		T :	TIME;
	END_VAR

	VAR_OUTPUT
		Y :	DWORD;
	END_VAR

	VAR
		last :	UDINT;
		tx :	UDINT;
		init :	BOOL;
		Yi :	REAL;
		T_PLC_MS :	T_PLC_MS_block;
	END_VAR

	T_PLC_MS();
	tx:= T_PLC_MS.T_PLC_MS;

	IF NOT init OR T = t#0s THEN
		init := TRUE;
		Yi := _DWORD_TO_REAL(X);
	ELSE
		Yi := Yi + (_DWORD_TO_REAL(X) - _DWORD_TO_REAL(Y)) * UDINT_TO_REAL(tx - last) / TIME_TO_REAL(T);
	END_IF;
	last := tx;

	Y := _REAL_TO_DWORD(Yi);

END_FUNCTION_BLOCK

PROGRAM program0
  VAR
	X :	DWORD;
	T :	TIME;

	Y :	DWORD;

	func_block : FILTER_DW;
  END_VAR
	func_block.X  := X;
	func_block.T  := T;
	func_block();
	Y := func_block.Y;
END_PROGRAM

CONFIGURATION Config0
	VAR_GLOBAL
		PLC_TICKS_PER_SEC :	INT;
		PLC_SYS_TICK_CNT :	DINT;
	END_VAR
	RESOURCE Res0 ON PLC
		TASK task0(INTERVAL := T#20ms,PRIORITY := 0);
		PROGRAM instance0 WITH task0 : program0;
	END_RESOURCE
END_CONFIGURATION

(* ---- FILTER_I.ST ---- *)
FUNCTION_BLOCK T_PLC_MS_block
	VAR_OUTPUT
		T_PLC_MS :	UDINT;
	END_VAR

	VAR_EXTERNAL
		PLC_TICKS_PER_SEC :	INT;
		PLC_SYS_TICK_CNT :	DINT;
	END_VAR

	VAR
		debug :	BOOL;(*Debug-Mode ON / OFF*)
		N :	INT;(*Debug-Faktor*)
		Offset :	UDINT;(*Debug-Offset*)
		temp :	DWORD := DWORD#1;(*Debug-Offset*)
		mode :	BOOL;(*modus*)
		faktor :	UDINT;(*Systemtakt-Faktor*)
		init :	BOOL;
		v_plc_ticks_per_sec :	UDINT;
		base :	UDINT := UDINT#1000;
	END_VAR

	IF init = FALSE THEN
		v_plc_ticks_per_sec := INT_TO_UDINT(PLC_TICKS_PER_SEC);
		IF v_plc_ticks_per_sec = UDINT#1024 THEN
			faktor := UDINT#1;
			mode := FALSE;
		ELSIF v_plc_ticks_per_sec > UDINT#0 THEN
			IF v_plc_ticks_per_sec <= base THEN
				faktor := base / v_plc_ticks_per_sec;
				mode := FALSE;
			ELSE
				faktor := v_plc_ticks_per_sec / base;
				mode := TRUE;
			END_IF;
		ELSE
			faktor := UDINT#1;
		END_IF;
		init := TRUE;
	END_IF;

	IF mode THEN
		T_PLC_MS := DINT_TO_UDINT(PLC_SYS_TICK_CNT) / faktor;
	ELSE
		T_PLC_MS := DINT_TO_UDINT(PLC_SYS_TICK_CNT) * faktor;
	END_IF;

	IF debug THEN
		T_PLC_MS := (DWORD_TO_UDINT(SHL(UDINT_TO_DWORD(T_PLC_MS),N) OR SHL(temp,N)) - UDINT#1) + Offset;
	END_IF;

END_FUNCTION_BLOCK

FUNCTION_BLOCK FILTER_I
	VAR_INPUT
		X :	INT;
		T :	TIME;
	END_VAR

	VAR_OUTPUT
		Y :	INT;
	END_VAR

	VAR
		Yi :	DINT;
		last :	UDINT;
		tx :	UDINT;
		init :	BOOL;
		T_PLC_MS :	T_PLC_MS_block;
	END_VAR

	T_PLC_MS();
	tx:= T_PLC_MS.T_PLC_MS;

	IF NOT init OR T = t#0s THEN
		init := TRUE;
		Yi := INT_TO_DINT(X) * DINT#1000;
	ELSE
		Yi := Yi + INT_TO_DINT(X - Y) * UDINT_TO_DINT(tx - last) * DINT#1000 / TIME_TO_DINT(T);
	END_IF;
	last := tx;
	Y := DINT_TO_INT(yi / DINT#1000);

END_FUNCTION_BLOCK

PROGRAM program0
  VAR
	X :	INT;
	T :	TIME;

	Y :	INT;

	func_block : FILTER_I;
  END_VAR
	func_block.X  := X;
	func_block.T  := T;
	func_block();
	Y := func_block.Y;
END_PROGRAM

CONFIGURATION Config0
	VAR_GLOBAL
		PLC_TICKS_PER_SEC :	INT;
		PLC_SYS_TICK_CNT :	DINT;
	END_VAR
	RESOURCE Res0 ON PLC
		TASK task0(INTERVAL := T#20ms,PRIORITY := 0);
		PROGRAM instance0 WITH task0 : program0;
	END_RESOURCE
END_CONFIGURATION

(* ---- FILTER_MAV_DW.ST ---- *)
TYPE
  oscat_ardw_0_31             : ARRAY [0..31]   OF DWORD;
END_TYPE

FUNCTION INC1:INT

	VAR_INPUT
		X :	INT;
		N :	INT;
	END_VAR

	IF X >= N - 1 THEN
		INC1 := 0;
	ELSE
		INC1 := X + 1;
	END_IF;
END_FUNCTION

FUNCTION_BLOCK FILTER_MAV_DW

	VAR_INPUT
		X :	DWORD;
		N :	UINT;
		RST :	BOOL;
	END_VAR

	VAR_OUTPUT
		Y :	DWORD;
	END_VAR

	VAR
		init :	BOOL;
		buffer :	oscat_ardw_0_31;
		i :	INT;
		tmp :	INT;
	END_VAR

	N := MIN(N, UINT#32);

	(* startup initialisation *)
	IF NOT init OR rst OR N = UINT#0 THEN
		init := TRUE;
		tmp := UINT_TO_INT(N)-1;
		FOR i := 0 TO tmp DO
			buffer[i] := X;
		END_FOR;
		Y := X;
	ELSE
		tmp := UINT_TO_INT(N);
		i := INC1(i, tmp);
		Y := UDINT_TO_DWORD(DWORD_TO_UDINT(Y) + (DWORD_TO_UDINT(X) - DWORD_TO_UDINT(buffer[i])) / UINT_TO_UDINT(N));
		buffer[i] := X;
	END_IF;

END_FUNCTION_BLOCK

PROGRAM program0
  VAR
	X :	DWORD;
	N :	UINT;
	RST :	BOOL;

	Y :	DWORD;

	func_block : FILTER_MAV_DW;
  END_VAR
	func_block.X  := X;
	func_block.N  := N;
	func_block.RST  := RST;
	func_block();
	Y := func_block.Y;
END_PROGRAM

CONFIGURATION Config0

	RESOURCE Res0 ON PLC
		TASK task0(INTERVAL := T#20ms,PRIORITY := 0);
		PROGRAM instance0 WITH task0 : program0;
	END_RESOURCE
END_CONFIGURATION

(* ---- FILTER_MAV_W.ST ---- *)
TYPE
  oscat_FILTER_MAV_W          : ARRAY [0..31]   OF WORD;
END_TYPE

FUNCTION INC1:INT

	VAR_INPUT
		X :	INT;
		N :	INT;
	END_VAR

	IF X >= N - 1 THEN
		INC1 := 0;
	ELSE
		INC1 := X + 1;
	END_IF;
END_FUNCTION

FUNCTION_BLOCK FILTER_MAV_W
	VAR_INPUT
		X :	WORD;
		N :	UINT;
		RST :	BOOL;
	END_VAR

	VAR_OUTPUT
		Y :	WORD;
	END_VAR

	VAR
		init :	BOOL;
		buffer :	oscat_FILTER_MAV_W;
		i :	INT;
		sum :	UDINT;
		tmp :	INT;
	END_VAR

	N := MIN(N, UINT#32);

	(* startup initialisation *)
	IF NOT init OR rst OR N = UINT#0 THEN
		init := TRUE;
		tmp := UINT_TO_INT(N) - 1;
		FOR i := 1 TO tmp DO
			buffer[i] := X;
		END_FOR;
		sum := UINT_TO_UDINT(WORD_TO_UINT(Y) * N);
		Y := X;
	ELSE
		tmp := UINT_TO_INT(N);
		i := INC1(i, tmp);
		sum := sum + WORD_TO_UDINT(X) - WORD_TO_UDINT(buffer[i]);
		Y := UDINT_TO_WORD(sum / UINT_TO_UDINT(N));
		buffer[i] := X;
	END_IF;

END_FUNCTION_BLOCK

PROGRAM program0
  VAR
	X :	WORD;
	N :	UINT;
	RST :	BOOL;

	Y :	WORD;

	func_block : FILTER_MAV_W;
  END_VAR
	func_block.X  := X;
	func_block.N  := N;
	func_block.RST  := RST;
	func_block();
	Y := func_block.Y;
END_PROGRAM

CONFIGURATION Config0

	RESOURCE Res0 ON PLC
		TASK task0(INTERVAL := T#20ms,PRIORITY := 0);
		PROGRAM instance0 WITH task0 : program0;
	END_RESOURCE
END_CONFIGURATION

(* ---- FILTER_W.ST ---- *)
FUNCTION_BLOCK T_PLC_MS_block
	VAR_OUTPUT
		T_PLC_MS :	UDINT;
	END_VAR

	VAR_EXTERNAL
		PLC_TICKS_PER_SEC :	INT;
		PLC_SYS_TICK_CNT :	DINT;
	END_VAR

	VAR
		debug :	BOOL;(*Debug-Mode ON / OFF*)
		N :	INT;(*Debug-Faktor*)
		Offset :	UDINT;(*Debug-Offset*)
		temp :	DWORD := DWORD#1;(*Debug-Offset*)
		mode :	BOOL;(*modus*)
		faktor :	UDINT;(*Systemtakt-Faktor*)
		init :	BOOL;
		v_plc_ticks_per_sec :	UDINT;
		base :	UDINT := UDINT#1000;
	END_VAR

	IF init = FALSE THEN
		v_plc_ticks_per_sec := INT_TO_UDINT(PLC_TICKS_PER_SEC);
		IF v_plc_ticks_per_sec = UDINT#1024 THEN
			faktor := UDINT#1;
			mode := FALSE;
		ELSIF v_plc_ticks_per_sec > UDINT#0 THEN
			IF v_plc_ticks_per_sec <= base THEN
				faktor := base / v_plc_ticks_per_sec;
				mode := FALSE;
			ELSE
				faktor := v_plc_ticks_per_sec / base;
				mode := TRUE;
			END_IF;
		ELSE
			faktor := UDINT#1;
		END_IF;
		init := TRUE;
	END_IF;

	IF mode THEN
		T_PLC_MS := DINT_TO_UDINT(PLC_SYS_TICK_CNT) / faktor;
	ELSE
		T_PLC_MS := DINT_TO_UDINT(PLC_SYS_TICK_CNT) * faktor;
	END_IF;

	IF debug THEN
		T_PLC_MS := (DWORD_TO_UDINT(SHL(UDINT_TO_DWORD(T_PLC_MS),N) OR SHL(temp,N)) - UDINT#1) + Offset;
	END_IF;

END_FUNCTION_BLOCK

FUNCTION_BLOCK FILTER_W
	VAR_INPUT
		X :	WORD;
		T :	TIME;
	END_VAR

	VAR_OUTPUT
		Y :	WORD;
	END_VAR

	VAR
		last :	UDINT;
		tx :	UDINT;
		init :	BOOL;
		tmp :	DINT;
		T_PLC_MS :	T_PLC_MS_Block;
	END_VAR

	T_PLC_MS();
	tx:= T_PLC_MS.T_PLC_MS;

	IF NOT init OR T = T#0s THEN
		init := TRUE;
		last := tx;
		Y := X;
	ELSIF Y = X THEN
		last := tx;
	ELSE
		tmp := UINT_TO_DINT(WORD_TO_UINT(X) - WORD_TO_UINT(Y)) * UDINT_TO_DINT(tx - last) / TIME_TO_DINT(T);
		IF tmp <> DINT#0 THEN
			Y := DINT_TO_WORD(WORD_TO_DINT(Y) + tmp);
			last := tx;
		END_IF;
	END_IF;

END_FUNCTION_BLOCK

PROGRAM program0
  VAR
	X :	WORD;
	T :	TIME;

	Y :	WORD;

	func_block : FILTER_W;
  END_VAR
	func_block.X  := X;
	func_block.T  := T;
	func_block();
	Y := func_block.Y;
END_PROGRAM

CONFIGURATION Config0
	VAR_GLOBAL
		PLC_TICKS_PER_SEC :	INT;
		PLC_SYS_TICK_CNT :	DINT;
	END_VAR
	RESOURCE Res0 ON PLC
		TASK task0(INTERVAL := T#20ms,PRIORITY := 0);
		PROGRAM instance0 WITH task0 : program0;
	END_RESOURCE
END_CONFIGURATION

(* ---- FILTER_WAV.ST ---- *)
TYPE
  oscat_arr_0_15              : ARRAY [0..15]   OF REAL;
END_TYPE

FUNCTION INC1:INT

	VAR_INPUT
		X :	INT;
		N :	INT;
	END_VAR

	IF X >= N - 1 THEN
		INC1 := 0;
	ELSE
		INC1 := X + 1;
	END_IF;
END_FUNCTION

FUNCTION DEC1:INT

	VAR_INPUT
		X :	INT;
		N :	INT;
	END_VAR

	IF X = 0 THEN
		DEC1 := N - 1;
	ELSE
		DEC1 := X - 1;
	END_IF;

END_FUNCTION

FUNCTION_BLOCK FILTER_WAV
	VAR_INPUT
		X :	REAL;
		W :	oscat_arr_0_15;
		RST :	BOOL;
	END_VAR

	VAR_OUTPUT
		Y :	REAL;
	END_VAR

	VAR
		init :	BOOL;
		buffer :	oscat_arr_0_15;
		i :	INT;
		n :	INT;
	END_VAR

	IF NOT init OR rst THEN
		init := TRUE;
		FOR i := 0 TO 15 DO
			buffer[i] := X;
		END_FOR;
		i := 15;
		Y := X;
	ELSE
		i := INC1(i, 16);
		buffer[i] := X;
	END_IF;

	Y := 0.0;
	FOR n := 0 TO 15 DO
		Y := buffer[i] * W[n] + Y;
		i := DEC1(i, 16);
	END_FOR;
END_FUNCTION_BLOCK

PROGRAM program0
  VAR
	X :	REAL;
	W :	oscat_arr_0_15;
	RST :	BOOL;

	Y :	REAL;

	func_block : FILTER_WAV;
  END_VAR
	func_block.X  := X;
	func_block.W  := W;
	func_block.RST  := RST;
	func_block();
	Y := func_block.Y;
END_PROGRAM

CONFIGURATION Config0

	RESOURCE Res0 ON PLC
		TASK task0(INTERVAL := T#20ms,PRIORITY := 0);
		PROGRAM instance0 WITH task0 : program0;
	END_RESOURCE
END_CONFIGURATION

(* ---- FINDB.ST ---- *)
FUNCTION_BLOCK FINDB_Block

	VAR_INPUT
		STR1 :	STRING;
		STR2 :	STRING;
	END_VAR

	VAR_OUTPUT
		FINDB :	INT;
	END_VAR

	VAR
		pos :	INT;
		length :	INT;
		string_temp :	STRING;
	END_VAR

	length := LEN(str2);
	pos := LEN(str1) - length +1;
	WHILE (pos >= 1) DO
		string_temp := MID(str1,length,pos);
		IF EQ_STRING(string_temp,str2) THEN
			FindB := pos;
			RETURN;
		END_IF;
	pos := pos -1;
	END_WHILE;
	FindB := 0;

END_FUNCTION_BLOCK

PROGRAM program0
  VAR
		STR1 :	STRING;
		STR2 :	STRING;

		FINDB :	INT;

	func_block : FINDB_Block;
  END_VAR
	func_block.STR1  := STR1;
	func_block.STR2  := STR2;
	func_block();
	FINDB := func_block.FINDB;
END_PROGRAM

CONFIGURATION Config0

	RESOURCE Res0 ON PLC
		TASK task0(INTERVAL := T#20ms,PRIORITY := 0);
		PROGRAM instance0 WITH task0 : program0;
	END_RESOURCE
END_CONFIGURATION

(* ---- FINDB_NONUM.ST ---- *)
FUNCTION_BLOCK FINDB_NONUM_Block

	VAR_INPUT
		STR :	STRING;
	END_VAR

	VAR_OUTPUT
		FINDB_NONUM :	INT;
	END_VAR

	VAR
		pos :	INT;
		x :	INT;
	END_VAR

	pos := LEN(str);
	WHILE (pos >=1) DO
		x :=GET_CHAR(str,pos);
		IF (X < 48 AND X <> 46) OR X > 57 THEN
			findB_nonum := pos;
			RETURN;
		END_IF;
	pos := pos -1;
	END_WHILE;
	findB_nonum := 0;

END_FUNCTION_BLOCK

PROGRAM program0
	VAR
		STR :	STRING;

		FINDB_NONUM :	INT;

		func_block : FINDB_NONUM_Block;
	END_VAR
	func_block.STR := STR;
	func_block();
	FINDB_NONUM  := func_block.FINDB_NONUM;
END_PROGRAM

CONFIGURATION Config0
	RESOURCE Res0 ON PLC
		TASK task0(INTERVAL := T#20ms,PRIORITY := 0);
		PROGRAM instance0 WITH task0 : program0;
	END_RESOURCE
END_CONFIGURATION

(* ---- FINDP.ST ---- *)
FUNCTION_BLOCK FINDP_Block

	VAR_INPUT
		STR :	STRING;
		SRC :	STRING;
		POS :	INT;
	END_VAR

	VAR_OUTPUT
		FINDP :	INT;
	END_VAR

	VAR
		i :	INT;
		ls :	INT;
		lx :	INT;
		stp :	INT;
		st_tmp :	STRING;
	END_VAR

	ls := LEN(str);
	lx := LEN(src);
	IF ls < lx OR lx = 0 THEN RETURN; END_IF;
	stp := ls - lx + 1;
	FOR i := MAX(pos,1) TO stp DO
		st_tmp := MID(str,lx,i);
		IF EQ_STRING(st_tmp,src) THEN
			FINDP := i;
			RETURN;
		END_IF;
	END_FOR;
	FINDP := 0;

END_FUNCTION_BLOCK

PROGRAM program0

	VAR
		STR :	STRING;
		SRC :	STRING;
		POS :	INT;

        FINDP :	INT;
		func_block : FINDP_Block;
	END_VAR
		func_block.STR := STR;
		func_block.SRC := SRC;
		func_block.POS := POS;
		func_block();
		FINDP := func_block.FINDP;

END_PROGRAM

CONFIGURATION Config0

	RESOURCE Res0 ON PLC
		TASK task0(INTERVAL := T#20ms,PRIORITY := 0);
		PROGRAM instance0 WITH task0 : program0;
	END_RESOURCE

END_CONFIGURATION

(* ---- FIX.ST ---- *)
FUNCTION _BYTE_TO_INT:INT
	VAR_INPUT
		IN :	BYTE;
	END_VAR

	_BYTE_TO_INT := USINT_TO_INT(BYTE_TO_USINT(IN));
END_FUNCTION

FUNCTION_BLOCK CHR_TO_STRING_Block
	VAR_INPUT
		C :	BYTE;
	END_VAR

	VAR_OUTPUT
		CHR_TO_STRING :	STRING;
	END_VAR

	CHR_TO_STRING := BYTE_TO_STRING(C);

END_FUNCTION_BLOCK

FUNCTION BIT_OF_DWORD : BOOL
  VAR_INPUT
    IN : DWORD;
    N : INT;
  END_VAR

  BIT_OF_DWORD := (SHR(in,N) AND 16#00000001) > 0;
  (* from OSCAT library; www.oscat.de  *)
END_FUNCTION

FUNCTION_BLOCK FILL_Block
	VAR_INPUT
		C :	BYTE;
		L :	INT;
	END_VAR

	VAR_OUTPUT
		FILL :	STRING;
	END_VAR

	VAR
		N :	BYTE;
		I :	INT;
		sx :	STRING;
		CHR_TO_STRING :	CHR_TO_STRING_Block;
		FILL_tmp :	STRING;
	END_VAR

	CHR_TO_STRING(C:=c);
	Sx:=CHR_TO_STRING.CHR_TO_STRING;
	(* create string *)
	N := INT_TO_BYTE(LIMIT(0,L,80));
	(* create a string of characters to be connected to str *)
	FILL := '';
	FOR i := 1 TO 8 DO
		FILL_tmp := FILL;
		FILL := CONCAT(FILL_tmp,FILL);
		IF BIT_OF_DWORD(BYTE_TO_DWORD(N),7) THEN FILL := CONCAT(FILL,Sx); END_IF;
		N := SHL(N,1);
	END_FOR;
END_FUNCTION_BLOCK

FUNCTION_BLOCK FIX_Block

	VAR_INPUT
		STR :	STRING;
		L :	INT;
		C :	BYTE;
		M :	INT;
	END_VAR

	VAR_OUTPUT
		FIX :	STRING;
	END_VAR

	VAR
		N :	INT;
		FILL :	FILL_Block;
	END_VAR

	N := LIMIT(0,L,255) - LEN(str);
	IF N <= 0 THEN
		(* truncate the string at length N *)
		IF M = 1 THEN
			FIX := RIGHT(str,L);
		ELSE
			FIX := LEFT(str,L);
		END_IF;
	ELSIF M = 1 THEN
		(* connect fill characters at the beginning *)
		FILL(C:=C,L:=N);
		FIX := CONCAT(FILL.FILL,str);
	ELSIF M = 2 THEN
		(* center str beween fill characters *)
		(* for an uneven number of fill characters, there is one more at the end *)
		FILL(C:=C,L:=_BYTE_TO_INT(SHR(INT_TO_BYTE(N+1),1)));
		FIX := CONCAT(str,FILL.FILL);
		FILL(C:=C,L:=_BYTE_TO_INT(SHR(INT_TO_BYTE(N),1)));
		FIX := CONCAT(FILL.FILL,FIX);
	ELSE
		(* connect fill characters at the end *)
		FILL(C:=C,L:=N);
		FIX := CONCAT(str,FILL.FILL);
	END_IF;

END_FUNCTION_BLOCK

PROGRAM program0
  VAR
	STR :	STRING;
	L   :	INT;
	C   :	BYTE;
	M   :	INT;

	FIX :	STRING;

	func_block : FIX_Block;
  END_VAR
	func_block.STR:=STR;
	func_block.L  :=L  ;
	func_block.C  :=C  ;
	func_block.M  :=M  ;
	func_block();
	FIX := func_block.FIX;
END_PROGRAM

CONFIGURATION Config0
  RESOURCE Res0 ON PLC
    TASK task0(INTERVAL := T#20ms,PRIORITY := 0);
    PROGRAM instance0 WITH task0 : program0;
  END_RESOURCE
END_CONFIGURATION
